(* IEC 61131-3 sources: daoli-st-library/DL_Process (part 54) *)

(* ---- FB_DL_SugarPanBatchSeq.st ---- *)
(*==============================================================================
  Component : FB_DL_SugarPanBatchSeq
  Category  : DL_Process
  Type      : FB
  Complexity: C4
  VERSION   : v1.0.0
  功能      : 煮糖罐批次时序（抽真空→进糖浆→浓缩→投晶种→助晶→终浓缩→破真空→放糖→洗罐）
  开源溯源  : 道莅原创 clean-room 自研（无外部代码引用）｜License: MIT
  边界条件  : ① 相迁移主判据为过饱和度 S（本件内联调用 CalcSupersaturation 计算）：
                 S = (Bx / (100 − Bx)) / (BxSat / (100 − BxSat))，BxSat = fSolA + fSolB × 温度；
                 该式为工程线性溶解度近似，精度受 fSolA / fSolB 标定限，不适用于高纯度精糖结晶建模。
              ② 真空与温度双联锁：真空丧失（fVacKpa 高于 fVacGoodKpa）或温度超上限 -> E3 立即断能；
                 温度低于下限 -> E2 停机待复位（糖液过冷会在罐内结块，属可恢复但需人工确认）。
              ③ 黄级语义：助晶相过饱和度超 fSWarn 只记录分级、不迁移、不置 bError（红/黑才动作）。
              ④ 过饱和度计算为「正解方向」：域外输入返回哨兵 0.0 并由调用方升 E2 上报（不静默钳位）。
                 S 物理上恒 > 1（过饱和），故 0.0 与任何合法值不重叠（R81 哨兵口径）。
                 传感器域判只在批次运行相生效——空闲相罐内空载（锤度 0、常压）属正常读数，不得误锁故障。
              ⑤ 默认引脚组合自证（R114）：握手类（bSyrupReady / bSeedAdded / bDischargeDone / bWashDone）
                 默认 FALSE，默认组合无法越过进料与放料握手直达完成相；使能类（bEStopHealthy）默认 TRUE
                 与 bEnable 同族，断线由硬件安全回路保证。
              ⑥ 复位作用域（R311）：bReset 沿清 E2/E3 锁存 + 批次计数 + 曲线锁存；bStop 只清 E2 与相位。
  状态机    : eIdle 待机 / eVacuum 抽真空 / eFillSyrup 进糖浆 / eConcentrate 浓缩到过饱和 /
              eSeed 投晶种 / eGrow 助晶养晶 / eFinalBoil 终浓缩到放糖锤度 / eBreakVac 破真空 /
              eDischarge 放糖 / eWash 洗罐 / eDone 结算拍 / eFault 停机待复位(E2) / eSafeStop 安全断能(E3)
  自检      : R1 零 GVL ｜ R2 零物理地址 ｜ R3 纯 IEC 61131-3 ｜ R4 除零先判 + 非有限自反判 ｜
              R6 CASE 含 ELSE ｜ R7 九 TON 两沿段 0 无条件刷新 ｜ R10 仅标准转换函数 ｜ R14 无属性件
==============================================================================*)
TYPE E_DL_SpbPhase :
(
    eIdle        := 0,  (* 待机：等启动沿 / Idle, waiting for start edge *)
    eVacuum      := 10, (* 抽真空相：真空度达标 / Pulling vacuum *)
    eFillSyrup   := 20, (* 进糖浆相：进料到量 / Filling syrup *)
    eConcentrate := 30, (* 浓缩相：S 到投晶目标 / Concentrating to seeding S *)
    eSeed        := 40, (* 投晶种相：晶种加入完成 / Seeding *)
    eGrow        := 50, (* 助晶相：养晶至目标 S / Crystal growing *)
    eFinalBoil   := 60, (* 终浓缩相：锤度到放糖点 / Final boil to discharge Brix *)
    eBreakVac    := 70, (* 破真空相：破真空到位 / Breaking vacuum *)
    eDischarge   := 80, (* 放糖相：放料完成 / Discharging *)
    eWash        := 90, (* 洗罐相：洗罐完成 / Pan washing *)
    eDone        := 100,(* 结算拍：批次与节拍统计 / Settlement, one-scan *)
    eFault       := 110,(* 停机待复位（E2）/ Stop awaiting reset, E2 *)
    eSafeStop    := 120 (* 安全侧断能（E3）/ Safety energy cut, E3 *)
);
END_TYPE
TYPE E_DL_SpbCause :
(
    eNone       := 0,   (* 无异常 / No anomaly *)
    eVacLost    := 1,   (* 真空度丧失（E3）/ Vacuum lost, E3 *)
    eTempHigh   := 2,   (* 罐温超上限（E3）/ Over-temperature, E3 *)
    eTempLow    := 3,   (* 罐温低于下限（E2，过冷结块）/ Under-temperature, E2 *)
    eSigBad     := 4,   (* 传感器非有限或 S 计算域外（E2）/ Non-finite signal or S out of domain, E2 *)
    eEStopOpen  := 5,   (* 急停回路断开（E3）/ E-stop open, E3 *)
    eVacTmo     := 6,   (* 抽真空超时（E2）/ Vacuum timeout, E2 *)
    eFillTmo    := 7,   (* 进糖浆超时（E2）/ Fill timeout, E2 *)
    eConcTmo    := 8,   (* 浓缩超时（E2）/ Concentrate timeout, E2 *)
    eSeedTmo    := 9,   (* 投晶种超时（E2）/ Seeding timeout, E2 *)
    eGrowTmo    := 10,  (* 助晶超时（E2）/ Growing timeout, E2 *)
    eFinalTmo   := 11,  (* 终浓缩超时（E2）/ Final boil timeout, E2 *)
    eBreakTmo   := 12,  (* 破真空超时（E2）/ Break-vacuum timeout, E2 *)
    eDischTmo   := 13,  (* 放糖超时（E2）/ Discharge timeout, E2 *)
    eWashTmo    := 14,  (* 洗罐超时（E2）/ Wash timeout, E2 *)
    eCfgBad     := 15,  (* 组态非法（E2）/ Illegal configuration, E2 *)
    ePhaseBad   := 16   (* 非法相位兜底（E2）/ Illegal phase fallback, E2 *)
);
END_TYPE
TYPE E_DL_SpbGrade :
(
    eOk     := 0,       (* 无异常 / No anomaly *)
    eYellow := 1,       (* 黄：记录并继续（S 偏离不升故障）/ Yellow, recorded only *)
    eRed    := 2,       (* 红：本批次降级（可继续至放糖）/ Red, batch degraded *)
    eBlack  := 3        (* 黑：立即断能 / Black, immediate energy cut *)
);
END_TYPE

FUNCTION_BLOCK FB_DL_SugarPanBatchSeq
VAR_INPUT
    bStart          : BOOL := FALSE;    (* 启动沿（eIdle 入 eVacuum） [-] / Start rising edge *)
    bStop           : BOOL := FALSE;    (* 中止：回 eIdle 并清 E2 锁存 [-] / Abort, clears E2 only *)
    bReset          : BOOL := FALSE;    (* 复位沿：清全部锁存 + 批次计数（R311） [-] / Reset edge *)
    bSyrupReady     : BOOL := FALSE;    (* 进糖浆到位（默认 FALSE 禁跳步） [-] / Syrup fill in position *)
    bSeedAdded      : BOOL := FALSE;    (* 晶种已加入（默认 FALSE 禁跳步） [-] / Seed added *)
    bDischargeDone  : BOOL := FALSE;    (* 放糖完成（默认 FALSE 禁跳步） [-] / Discharge done *)
    bWashDone       : BOOL := FALSE;    (* 洗罐完成（默认 FALSE 禁跳步） [-] / Wash done *)
    bEStopHealthy   : BOOL := TRUE;     (* 急停回路正常（使能类引脚，默认 TRUE） [-] / E-stop healthy *)
    fVacKpa         : LREAL := 101.3;   (* 罐内绝对压力实测（真空好 = 值低） [kPa] / Pan absolute pressure [kPa] *)
    fTempC          : LREAL := 20.0;    (* 糖液温度实测 [℃] / Syrup temperature [degC] *)
    fBrix           : LREAL := 65.0;    (* 糖液锤度实测，域 0..100 [°Bx] / Brix [degBx] *)
    fVacGoodKpa     : LREAL := 30.0;    (* 真空良好门限，域 > 0（实测 <= 该值即真空有效） [kPa] / Vacuum good limit [kPa] *)
    fTempMinC       : LREAL := 60.0;    (* 罐温下限，域 > 0（低于则 E2） [℃] / Temperature floor [degC] *)
    fTempMaxC       : LREAL := 80.0;    (* 罐温上限，域 > fTempMinC（高于则 E3） [℃] / Temperature ceiling [degC] *)
    fSolA           : LREAL := 60.0;    (* 溶解度线性式截距（标定值），域 > 0 [°Bx] / Solubility intercept [degBx] *)
    fSolB           : LREAL := 0.25;    (* 溶解度线性式斜率（标定值），域 > 0 [°Bx/℃] / Solubility slope [degBx/degC] *)
    fSSeed          : LREAL := 1.20;    (* 投晶目标过饱和度，域 > 1.0 [-] / Seeding supersaturation *)
    fSGrow          : LREAL := 1.35;    (* 助晶终点过饱和度，域 > fSSeed [-] / Growing end supersaturation *)
    fSWarn          : LREAL := 1.45;    (* 过饱和预警上界，域 > fSGrow（黄级记录） [-] / Supersaturation warn limit *)
    fBrixDischarge  : LREAL := 92.0;    (* 放糖锤度，域 0..100（且 > fBrix） [°Bx] / Discharge Brix [degBx] *)
    atPhaseTmo      : ARRAY[0..8] OF TIME := [T#20M, T#30M, T#120M, T#10M, T#240M, T#120M, T#10M, T#20M, T#30M];   (* 超时窗 [ms]，下标 0..8 = 抽真空/进料/浓缩/投晶/助晶/终浓/破真空/放糖/洗罐 / Phase windows [ms] *)
    fCycleSec       : LREAL := 0.0;     (* 扫描周期（<=0 用缺省 0.01s） [s] / Scan cycle [s] *)
END_VAR
VAR_OUTPUT
    eState          : E_DL_SpbPhase;    (* 当前相（HMI 诊断） [-] / Present phase *)
    eCause          : E_DL_SpbCause;    (* 成因（锁存回放，R189） [-] / Latched cause playback *)
    eGrade          : E_DL_SpbGrade;    (* 分级出口 [-] / Grade outlet *)
    bError          : BOOL;             (* 故障标志（E2/E3 为 TRUE） [-] / Error flag *)
    bSafeCut        : BOOL;             (* 安全侧断能指令（E3 常 TRUE 至复位） [-] / Safety energy cut *)
    bDone           : BOOL;             (* 单拍结算脉冲 [-] / One-scan done pulse *)
    bBoilActive     : BOOL;             (* 浓缩段指示（供 IO 层驱动蒸汽阀） [-] / Boiling indicator *)
    nBatchCount     : UDINT;            (* 累计批次数（饱和） [批] / Batch count, saturating *)
    fSLast          : LREAL;            (* 最近过饱和度（0 = 无效）/ 哨兵值与合法域不重叠 [-] / Last supersaturation *)
    fBrixLast       : LREAL;            (* 最近锤度 [°Bx] / Last Brix [degBx] *)
    tBatchLast      : TIME;             (* 最近一批总时长 [ms] / Last batch duration [ms] *)
END_VAR
VAR
    _ePhase      : E_DL_SpbPhase := E_DL_SpbPhase.eIdle;     (* 内部相（CASE 唯一写入目标） [-] / Internal phase *)
    _eCause      : E_DL_SpbCause := E_DL_SpbCause.eNone;     (* 成因锁存量 [-] / Latched cause *)
    _eGrade      : E_DL_SpbGrade := E_DL_SpbGrade.eOk;       (* 分级锁存量 [-] / Latched grade *)
    _bFault      : BOOL := FALSE;       (* E2 锁存位（解除 = bReset 沿或 bStop） [-] / E2 latch *)
    _bSafeLatch  : BOOL := FALSE;       (* E3 锁存位（解除 = bReset 沿且安全恢复） [-] / E3 latch *)
    _bFaultReq   : BOOL := FALSE;       (* 单拍 E2 请求（段 1 预清，段 6 落地） [-] / One-scan E2 request *)
    _bSafeReq    : BOOL := FALSE;       (* 单拍 E3 请求（段 1 预清，段 6 落地） [-] / One-scan E3 request *)
    _bDonePulse  : BOOL := FALSE;       (* 单拍结算标志（段 1 预清） [-] / One-scan done flag *)
    _bVacOk      : BOOL := FALSE;       (* 真空有效判据 [-] / Vacuum valid *)
    _bTempHigh   : BOOL := FALSE;       (* 罐温超上限当拍量 [-] / Over-temperature this scan *)
    _bTempLow    : BOOL := FALSE;       (* 罐温低于下限当拍量 [-] / Under-temperature this scan *)
    _bVacBad     : BOOL := FALSE;       (* 真空传感器非有限当拍量 [-] / Vacuum non-finite *)
    _bTempBad    : BOOL := FALSE;       (* 温度传感器非有限当拍量 [-] / Temperature non-finite *)
    _bBrixBad    : BOOL := FALSE;       (* 锤度非有限或域外当拍量 [-] / Brix non-finite or out of domain *)
    _bCfgBad     : BOOL := FALSE;       (* 组态非法当拍量 [-] / Configuration bad *)
    _fS          : LREAL := 0.0;        (* 当拍过饱和度（0 = 计算无效哨兵） [-] / Supersaturation this scan *)
    _fMsTmp      : LREAL := 0.0;        (* 批次时长毫秒暂存（转换前钳位） [ms] / Batch milliseconds scratch *)
    _bVacRequired: BOOL := FALSE;       (* 本相要求真空有效（进料至终浓缩）/ Vacuum required in phase *)
    _bBatchActive: BOOL := FALSE;       (* 批次运行相（空闲与故障相不计信号域判）/ Batch active phase *)
    _bSafeOk     : BOOL := FALSE;       (* 安全条件已恢复（E3 解除判据）/ Safety conditions recovered *)
    _fBrixLatch  : LREAL := 0.0;        (* 锤度锁存（出口留影） [°Bx] / Brix latch *)
    _fBatchAccS  : LREAL := 0.0;        (* 本批时长累加 [s] / Batch time accumulator *)
    _tBatchLast  : TIME := T#0S;        (* 最近批时长锁存 [ms] / Last batch duration latch *)
    _fCy         : LREAL := 0.0;        (* 当拍有效周期 [s] / Effective cycle *)
    _nBatch      : UDINT := 0;          (* 批次累计锁存（饱和） [批] / Batch count latch *)
    _nIdxChk     : INT := 0;            (* 相窗遍历索引（循环变量） [-] / Loop index *)
    tonVacuum    : TON;                 (* 抽真空超时（段 0 无条件调用） / Vacuum timeout *)
    tonFill      : TON;                 (* 进糖浆超时 / Fill timeout *)
    tonConcentrate: TON;                (* 浓缩超时 / Concentrate timeout *)
    tonSeed      : TON;                 (* 投晶种超时 / Seeding timeout *)
    tonGrow      : TON;                 (* 助晶超时 / Growing timeout *)
    tonFinalBoil : TON;                 (* 终浓缩超时 / Final boil timeout *)
    tonBreakVac  : TON;                 (* 破真空超时 / Break-vacuum timeout *)
    tonDischarge : TON;                 (* 放糖超时 / Discharge timeout *)
    tonWash      : TON;                 (* 洗罐超时 / Wash timeout *)
    rtStart      : R_TRIG;              (* 启动沿（段 0 无条件调用） / Start edge *)
    rtReset      : R_TRIG;              (* 复位沿（段 0 无条件调用） / Reset edge *)
END_VAR
VAR CONSTANT
    DL_SPB_CYDEF   : LREAL := 0.01;         (* 缺省扫描周期 [s] / Default scan cycle [s] *)
    DL_SPB_BRIXTOP : LREAL := 100.0;        (* 锤度与溶解度共用上界 [°Bx] / Brix and solubility ceiling *)
    DL_SPB_DENMIN  : LREAL := 1.0E-6;       (* 除法分母下限（判零） [-] / Divisor floor *)
    DL_SPB_BATMAX  : UDINT := 4294967295;   (* 批次计数饱和上限 [批] / Batch count ceiling *)
END_VAR

(*-----------------------------------------------------------------------------
  方法 CalcSupersaturation：过饱和度计算（正解方向，域闸四段式）
  四段：① 返回值预置哨兵 0.0 ② 域闸命中直接 RETURN（非有限 / 锤度域外 / 溶解度域外）
        ③ 域内才做两次除法（分母均已证明 > DL_SPB_DENMIN） ④ 结果非有限复检兜底
  契约：返回 0.0 = 计算无效（哨兵），S 物理恒 > 1，调用方据 0.0 升 E2 上报（禁静默钳位）。
-----------------------------------------------------------------------------*)
METHOD PUBLIC CalcSupersaturation : LREAL
VAR_INPUT
    fBrixIn  : LREAL := 0.0;    (* 锤度输入，域 (0, 100) [°Bx] / Brix input *)
    fTempIn  : LREAL := 0.0;    (* 温度输入 [℃] / Temperature input *)
    fSolAIn  : LREAL := 0.0;    (* 溶解度截距，域 > 0 [°Bx] / Solubility intercept *)
    fSolBIn  : LREAL := 0.0;    (* 溶解度斜率，域 > 0 [°Bx/℃] / Solubility slope *)
END_VAR
VAR
    fBxSat : LREAL := 0.0;      (* 该温度下饱和锤度 [°Bx] / Saturated Brix at temperature *)
    fNum   : LREAL := 0.0;      (* 分子 Bx / (100 − Bx) [-] / Numerator *)
    fDen   : LREAL := 0.0;      (* 分母 BxSat / (100 − BxSat) [-] / Denominator *)
    fS     : LREAL := 0.0;      (* 过饱和度暂存 [-] / Supersaturation scratch *)
END_VAR

CalcSupersaturation := 0.0;     (* ① 预置哨兵 / Preset sentinel *)
IF (fBrixIn <> fBrixIn) OR ((fBrixIn - fBrixIn) <> (fBrixIn - fBrixIn)) THEN
    CalcSupersaturation := 0.0; (* ② 锤度非有限 / Brix non-finite *)
    RETURN;
END_IF
IF (fTempIn <> fTempIn) OR ((fTempIn - fTempIn) <> (fTempIn - fTempIn)) THEN
    CalcSupersaturation := 0.0; (* ② 温度非有限 / Temperature non-finite *)
    RETURN;
END_IF
IF (fSolAIn <= 0.0) OR (fSolBIn <= 0.0) THEN
    CalcSupersaturation := 0.0; (* ② 溶解度系数域外 / Solubility coefficient out of domain *)
    RETURN;
END_IF
IF (fBrixIn <= 0.0) OR (fBrixIn >= DL_SPB_BRIXTOP) THEN
    CalcSupersaturation := 0.0; (* ② 锤度域外（分母 100 − Bx 失效保护）/ Brix out of domain *)
    RETURN;
END_IF
fBxSat := fSolAIn + fSolBIn * fTempIn;                         (* 线性溶解度式 [°Bx] / Linear solubility *)
IF (fBxSat <= 0.0) OR (fBxSat >= DL_SPB_BRIXTOP) THEN
    CalcSupersaturation := 0.0; (* ② 饱和锤度域外 / Saturated Brix out of domain *)
    RETURN;
END_IF
fNum := fBrixIn / (DL_SPB_BRIXTOP - fBrixIn);                   (* ③ 分母 > 0 已证 / Denominator proven positive *)
fDen := fBxSat / (DL_SPB_BRIXTOP - fBxSat);                     (* ③ 分母 > 0 已证 / Denominator proven positive *)
IF fDen < DL_SPB_DENMIN THEN
    CalcSupersaturation := 0.0; (* ③ 分母判零（防御式，域闸后不可达）/ Divisor guard *)
    RETURN;
END_IF
fS := fNum / fDen;                                             (* 过饱和度 [-] / Supersaturation *)
IF (fS <> fS) OR ((fS - fS) <> (fS - fS)) THEN
    CalcSupersaturation := 0.0; (* ④ 结果非有限兜底 / Result non-finite fallback *)
    RETURN;
END_IF
CalcSupersaturation := fS;                                     (* 合法结果输出 / Valid result *)
END_METHOD

(*-----------------------------------------------------------------------------
  方法 ResetBatch：批次锁存复位（不清累计批次数，累计量只能由 bReset 沿清除）
  契约：返回 TRUE 表示复位执行；作用于分级、成因、过饱和度锁存与批次时长累加。
-----------------------------------------------------------------------------*)
METHOD PUBLIC ResetBatch : BOOL
ResetBatch := FALSE;                            (* 预置 / Preset *)
_eGrade := E_DL_SpbGrade.eOk;                   (* 清分级 / Clear grade *)
_eCause := E_DL_SpbCause.eNone;                 (* 清成因 / Clear cause *)
_fS := 0.0;                                     (* 清过饱和度哨兵 / Clear supersaturation *)
_fBrixLatch := 0.0;                             (* 清锤度锁存 / Clear Brix latch *)
_fBatchAccS := 0.0;                             (* 清批次时长累加 / Clear batch accumulator *)
ResetBatch := TRUE;                             (* 复位已执行 / Reset performed *)
END_METHOD

(* —— 段 0：传感器非有限与域判 + 过饱和度计算 + 组态闸 + 周期 + 九 TON 两沿无条件刷新（R7） —— *)
_bVacBad := (fVacKpa <> fVacKpa) OR ((fVacKpa - fVacKpa) <> (fVacKpa - fVacKpa));      (* NaN 自反 + Inf 差值 / NaN and Inf *)
_bTempBad := (fTempC <> fTempC) OR ((fTempC - fTempC) <> (fTempC - fTempC));
_bBrixBad := (fBrix <> fBrix) OR ((fBrix - fBrix) <> (fBrix - fBrix))
          OR (fBrix <= 0.0) OR (fBrix >= DL_SPB_BRIXTOP);                             (* 锤度域外并入信号级 / Brix domain *)
_bVacOk := (NOT _bVacBad) AND (fVacKpa <= fVacGoodKpa);                                (* 真空有效（值低为好）/ Vacuum valid *)
_bTempHigh := (NOT _bTempBad) AND (fTempC > fTempMaxC);                                (* 超上限（E3）/ Over-temperature *)
_bTempLow := (NOT _bTempBad) AND (fTempC < fTempMinC);                                 (* 低于下限（E2）/ Under-temperature *)
_fS := CalcSupersaturation(fBrix, fTempC, fSolA, fSolB);                               (* 过饱和度内联计算 / Supersaturation *)
_bCfgBad := (fVacGoodKpa <= 0.0) OR (fTempMinC <= 0.0) OR (fTempMaxC <= fTempMinC)
         OR (fSolA <= 0.0) OR (fSolB <= 0.0) OR (fBrixDischarge <= 0.0)
         OR (fBrixDischarge >= DL_SPB_BRIXTOP) OR (fSSeed <= 1.0)
         OR (fSGrow <= fSSeed) OR (fSWarn <= fSGrow);                                 (* 组态域闸与配比 / Config gate *)
FOR _nIdxChk := 0 TO 8 DO
    IF atPhaseTmo[_nIdxChk] <= T#0S THEN
        _bCfgBad := TRUE;                                                             (* 任一相窗非正 -> 组态非法 / Non-positive window *)
    END_IF
END_FOR
IF fCycleSec > 0.0 THEN
    _fCy := fCycleSec;                                                                (* 组态周期有效 / Configured cycle *)
ELSE
    _fCy := DL_SPB_CYDEF;                                                             (* 周期缺省兜底 / Default cycle *)
END_IF
rtStart(CLK := bStart);                                                               (* 启动沿，每拍必调 / Start edge every scan *)
rtReset(CLK := bReset);                                                               (* 复位沿，每拍必调 / Reset edge every scan *)
tonVacuum(IN := (_ePhase = E_DL_SpbPhase.eVacuum), PT := atPhaseTmo[0]);              (* 抽真空窗 / Vacuum window *)
tonFill(IN := (_ePhase = E_DL_SpbPhase.eFillSyrup), PT := atPhaseTmo[1]);             (* 进料窗 / Fill window *)
tonConcentrate(IN := (_ePhase = E_DL_SpbPhase.eConcentrate), PT := atPhaseTmo[2]);    (* 浓缩窗 / Concentrate window *)
tonSeed(IN := (_ePhase = E_DL_SpbPhase.eSeed), PT := atPhaseTmo[3]);                  (* 投晶窗 / Seeding window *)
tonGrow(IN := (_ePhase = E_DL_SpbPhase.eGrow), PT := atPhaseTmo[4]);                  (* 助晶窗 / Growing window *)
tonFinalBoil(IN := (_ePhase = E_DL_SpbPhase.eFinalBoil), PT := atPhaseTmo[5]);        (* 终浓窗 / Final boil window *)
tonBreakVac(IN := (_ePhase = E_DL_SpbPhase.eBreakVac), PT := atPhaseTmo[6]);          (* 破真空窗 / Break vacuum window *)
tonDischarge(IN := (_ePhase = E_DL_SpbPhase.eDischarge), PT := atPhaseTmo[7]);        (* 放糖窗 / Discharge window *)
tonWash(IN := (_ePhase = E_DL_SpbPhase.eWash), PT := atPhaseTmo[8]);                  (* 洗罐窗 / Wash window *)

(* —— 段 1：单拍量预清零（不含锁存/累加/计数，R107）+ 批次时长累加 —— *)
_bFaultReq := FALSE;                                                                  (* E2 请求预清 / E2 request preset *)
_bSafeReq := FALSE;                                                                   (* E3 请求预清 / E3 request preset *)
_bDonePulse := FALSE;                                                                 (* 结算标志预清 / Done preset *)
bError := FALSE;                                                                      (* 故障标志预清（出口汇总）/ Error preset *)
IF (_ePhase <> E_DL_SpbPhase.eIdle) AND (_ePhase <> E_DL_SpbPhase.eFault)
   AND (_ePhase <> E_DL_SpbPhase.eSafeStop) THEN
    _fBatchAccS := _fBatchAccS + _fCy;                                                (* 批次时长累加（仅工作相）/ Batch time, working phases only *)
END_IF
_bVacRequired := (_ePhase = E_DL_SpbPhase.eFillSyrup) OR (_ePhase = E_DL_SpbPhase.eConcentrate)
              OR (_ePhase = E_DL_SpbPhase.eSeed) OR (_ePhase = E_DL_SpbPhase.eGrow)
              OR (_ePhase = E_DL_SpbPhase.eFinalBoil);                                (* 真空维持段（放糖与洗罐不要求）/ Vacuum-required phases *)
_bBatchActive := (_ePhase <> E_DL_SpbPhase.eIdle) AND (_ePhase <> E_DL_SpbPhase.eDone)
                   AND (_ePhase <> E_DL_SpbPhase.eVacuum) AND (_ePhase <> E_DL_SpbPhase.eFillSyrup)   (* 空罐与进料相锤度天然为 0，不计入信号域判 / Exclude vacuum & fill phases: brix is naturally 0 *)
              AND (_ePhase <> E_DL_SpbPhase.eFault) AND (_ePhase <> E_DL_SpbPhase.eSafeStop);   (* 批次运行相判据 / Batch-active judge *)
_bSafeOk := bEStopHealthy AND (NOT _bTempHigh) AND (NOT _bTempBad);                   (* 安全恢复基础判据 / Base safety recovery *)
IF _eCause = E_DL_SpbCause.eVacLost THEN
    _bSafeOk := _bSafeOk AND _bVacOk;                                                 (* 真空成因须真空恢复（R152 可达性）/ Vacuum cause needs vacuum back *)
END_IF

(* —— 段 2：E3 安全侧（急停 / 真空丧失 / 罐温超上限）——最高优先级 —— *)
IF NOT bEStopHealthy THEN
    IF NOT _bSafeLatch THEN
        _bSafeReq := TRUE;                                                            (* 落地于段 6 / Landed in segment 6 *)
        _eCause := E_DL_SpbCause.eEStopOpen;                                          (* 归因：急停断开 / Cause: E-stop *)
    END_IF
ELSIF _bTempHigh THEN
    IF NOT _bSafeLatch THEN
        _bSafeReq := TRUE;
        _eCause := E_DL_SpbCause.eTempHigh;                                           (* 归因：超温 / Cause: over-temperature *)
    END_IF
ELSIF _bVacRequired AND (NOT _bVacBad) AND (NOT _bVacOk) THEN
    IF NOT _bSafeLatch THEN
        _bSafeReq := TRUE;                                                            (* 真空在非抽真空相丧失：立即断能 / Vacuum lost mid-batch *)
        _eCause := E_DL_SpbCause.eVacLost;                                            (* 归因：真空丧失 / Cause: vacuum lost *)
    END_IF
END_IF

(* —— 段 3：信号域闸与组态闸入 E2（E3 优先，安全相内不重复置因） —— *)
IF _bCfgBad AND (NOT _bSafeLatch) AND (NOT _bFault) THEN
    _bFaultReq := TRUE;                                                               (* 落地于段 6 / Landed in segment 6 *)
    _eCause := E_DL_SpbCause.eCfgBad;                                                 (* 归因：组态非法 / Cause: config *)
ELSIF _bBatchActive AND (_bVacBad OR _bBrixBad) THEN
    IF NOT _bSafeLatch AND NOT _bFault THEN
        _bFaultReq := TRUE;
        _eCause := E_DL_SpbCause.eSigBad;                                             (* 归因：传感器非有限 / Cause: non-finite *)
    END_IF
ELSIF _bBatchActive AND _bTempLow THEN
    IF NOT _bSafeLatch AND NOT _bFault THEN
        _bFaultReq := TRUE;
        _eCause := E_DL_SpbCause.eTempLow;                                            (* 归因：过冷 / Cause: under-temperature *)
    END_IF
ELSIF _bBatchActive AND (_fS <= 0.0) AND (NOT _bFault) THEN
    IF NOT _bSafeLatch THEN
        _bFaultReq := TRUE;                                                           (* S 计算域外（哨兵 0.0）/ S sentinel zero *)
        _eCause := E_DL_SpbCause.eSigBad;                                             (* 归因：S 计算域外 / Cause: S out of domain *)
    END_IF
END_IF

(* —— 段 4：迁出链（复位沿 > 中止；作用域逐项声明 R311） —— *)
IF rtReset.Q THEN
    _bFault := FALSE;                                                                 (* 作用域①：清 E2 锁存 / Clear E2 *)
    IF _bSafeOk THEN
        _bSafeLatch := FALSE;                                                         (* 作用域②：安全恢复才清 E3（成因相关判据）/ Clear E3 only if safe *)
    END_IF
    _eCause := E_DL_SpbCause.eNone;                                                   (* 作用域③：清成因分级 / Clear cause and grade *)
    _eGrade := E_DL_SpbGrade.eOk;
    _fS := 0.0;                                                                       (* 作用域④：清过饱和度锁存 / Clear supersaturation *)
    _fBrixLatch := 0.0;
    _fBatchAccS := 0.0;                                                               (* 作用域⑤：清批次时长 / Clear batch time *)
    _nBatch := 0;                                                                     (* 作用域⑥：清批次计数（生产资料复位）/ Clear batch count *)
    IF NOT _bSafeLatch THEN
        IF (_ePhase = E_DL_SpbPhase.eFault) OR (_ePhase = E_DL_SpbPhase.eSafeStop) THEN
            _ePhase := E_DL_SpbPhase.eIdle;                                           (* 作用域⑦：故障相迁回待机 / Back to idle *)
        END_IF
    END_IF
ELSIF bStop AND (_ePhase <> E_DL_SpbPhase.eIdle) AND (_ePhase <> E_DL_SpbPhase.eSafeStop) THEN
    IF _ePhase = E_DL_SpbPhase.eFault THEN
        _bFault := FALSE;                                                             (* 中止清 E2（E3 只由复位清）/ Abort clears E2 only *)
        _eCause := E_DL_SpbCause.eNone;
        _eGrade := E_DL_SpbGrade.eOk;
    END_IF
    _fBatchAccS := 0.0;                                                               (* 批次时长作废 / Batch time void *)
    _ePhase := E_DL_SpbPhase.eIdle;                                                   (* 回待机 / Back to idle *)
END_IF

(* —— 段 5：主状态机（过饱和度 / 锤度为相迁移主判据，超时为保护） —— *)
CASE _ePhase OF
E_DL_SpbPhase.eIdle:
    IF rtStart.Q AND (NOT _bFault) AND (NOT _bSafeLatch) THEN
        _eGrade := E_DL_SpbGrade.eOk;                                                 (* 新批起算 / New batch *)
        _eCause := E_DL_SpbCause.eNone;
        _fBatchAccS := 0.0;
        _ePhase := E_DL_SpbPhase.eVacuum;                                             (* 入抽真空相 / To vacuum *)
    END_IF
E_DL_SpbPhase.eVacuum:
    IF _bVacOk THEN
        _ePhase := E_DL_SpbPhase.eFillSyrup;                                          (* 真空达标 -> 进糖浆 / Vacuum OK, fill *)
    ELSIF tonVacuum.Q THEN
        _eCause := E_DL_SpbCause.eVacTmo;                                             (* 归因：抽真空超时 / Cause: vacuum timeout *)
        _bFaultReq := TRUE;
    END_IF
E_DL_SpbPhase.eFillSyrup:
    IF bSyrupReady THEN
        _ePhase := E_DL_SpbPhase.eConcentrate;                                        (* 进料到量 -> 浓缩 / Filled, concentrate *)
    ELSIF tonFill.Q THEN
        _eCause := E_DL_SpbCause.eFillTmo;                                            (* 归因：进料超时 / Cause: fill timeout *)
        _bFaultReq := TRUE;
    END_IF
E_DL_SpbPhase.eConcentrate:
    IF (_fS > 0.0) AND (_fS >= fSSeed) THEN
        _ePhase := E_DL_SpbPhase.eSeed;                                               (* S 到投晶目标 -> 投晶 / S reached, seed *)
    ELSIF tonConcentrate.Q THEN
        _eCause := E_DL_SpbCause.eConcTmo;                                            (* 归因：浓缩超时（S 未达）/ Cause: concentrate timeout *)
        _bFaultReq := TRUE;
    END_IF
E_DL_SpbPhase.eSeed:
    IF bSeedAdded THEN
        _ePhase := E_DL_SpbPhase.eGrow;                                               (* 晶种加入 -> 助晶 / Seeded, grow *)
    ELSIF tonSeed.Q THEN
        _eCause := E_DL_SpbCause.eSeedTmo;                                            (* 归因：投晶超时 / Cause: seeding timeout *)
        _bFaultReq := TRUE;
    END_IF
E_DL_SpbPhase.eGrow:
    IF (_fS > 0.0) AND (_fS > fSWarn) THEN
        _eGrade := E_DL_SpbGrade.eYellow;                                             (* 过饱和偏高预警（黄，只记录不迁移）/ High-S warning, recorded only *)
    END_IF
    IF (_fS > 0.0) AND (_fS >= fSGrow) THEN
        _ePhase := E_DL_SpbPhase.eFinalBoil;                                          (* 养晶到位 -> 终浓 / Grown, final boil *)
    ELSIF tonGrow.Q THEN
        _eCause := E_DL_SpbCause.eGrowTmo;                                            (* 归因：助晶超时 / Cause: growing timeout *)
        _bFaultReq := TRUE;
    END_IF
E_DL_SpbPhase.eFinalBoil:
    IF (NOT _bBrixBad) AND (fBrix >= fBrixDischarge) THEN
        _fBrixLatch := fBrix;                                                         (* 放糖锤度锁存 / Latch discharge Brix *)
        _ePhase := E_DL_SpbPhase.eBreakVac;                                           (* 锤度到量 -> 破真空 / Brix reached, break vacuum *)
    ELSIF tonFinalBoil.Q THEN
        _eCause := E_DL_SpbCause.eFinalTmo;                                           (* 归因：终浓超时（锤度未达）/ Cause: final boil timeout *)
        _bFaultReq := TRUE;
    END_IF
E_DL_SpbPhase.eBreakVac:
    IF (NOT _bVacBad) AND (fVacKpa >= fVacGoodKpa) THEN
        _ePhase := E_DL_SpbPhase.eDischarge;                                          (* 真空破除到位 -> 放糖（本拍事件优先，R275）/ Vacuum broken, discharge *)
    ELSIF tonBreakVac.Q THEN
        _eCause := E_DL_SpbCause.eBreakTmo;                                           (* 归因：破真空超时 / Cause: break-vacuum timeout *)
        _bFaultReq := TRUE;
    END_IF
E_DL_SpbPhase.eDischarge:
    IF bDischargeDone THEN
        _ePhase := E_DL_SpbPhase.eWash;                                               (* 放糖完成 -> 洗罐 / Discharged, wash *)
    ELSIF tonDischarge.Q THEN
        _eCause := E_DL_SpbCause.eDischTmo;                                           (* 归因：放糖超时 / Cause: discharge timeout *)
        _bFaultReq := TRUE;
    END_IF
E_DL_SpbPhase.eWash:
    IF bWashDone THEN
        _ePhase := E_DL_SpbPhase.eDone;                                               (* 洗罐完成 -> 结算 / Washed, settle *)
    ELSIF tonWash.Q THEN
        _eCause := E_DL_SpbCause.eWashTmo;                                            (* 归因：洗罐超时 / Cause: wash timeout *)
        _bFaultReq := TRUE;
    END_IF
E_DL_SpbPhase.eDone:
    _bDonePulse := TRUE;                                                              (* 单拍结算（段 1 预清）/ One-scan done *)
    _fMsTmp := _fBatchAccS * 1000.0;                                                  (* 秒 -> 毫秒 [ms] / Second to millisecond *)
    IF _fMsTmp > 2147483647.0 THEN
        _fMsTmp := 2147483647.0;                                                      (* 取整前实数上限兜底（R153）/ Real ceiling before truncation *)
    END_IF
    _tBatchLast := DINT_TO_TIME(LREAL_TO_DINT(_fMsTmp));                              (* 批次时长换算 / Batch duration *)
    _fBatchAccS := 0.0;                                                               (* 累加清零 / Clear accumulator *)
    IF _nBatch < DL_SPB_BATMAX THEN
        _nBatch := _nBatch + 1;                                                       (* 批次推进（容量载体判上限）/ Saturating batch count *)
    END_IF
    _ePhase := E_DL_SpbPhase.eIdle;                                                   (* 回待机 / Back to idle *)
E_DL_SpbPhase.eFault:
    bError := TRUE;                                                                   (* 故障相驻留（锁存回放）/ Fault residency *)
E_DL_SpbPhase.eSafeStop:
    bError := TRUE;                                                                   (* 安全相驻留（锁存回放）/ Safety residency *)
ELSE
    _eCause := E_DL_SpbCause.ePhaseBad;                                               (* 非法相位兜底 / Illegal phase fallback *)
    _bFaultReq := TRUE;                                                               (* 由段 6 落地 / Landed in segment 6 *)
END_CASE

(* —— 段 6：E2/E3 请求统一落地（分支内只写成因与请求，落地仅此一处，R187/R252） —— *)
IF _bSafeReq AND (NOT _bSafeLatch) THEN
    _bSafeLatch := TRUE;                                                              (* E3 锁存 / Latch E3 *)
    _eGrade := E_DL_SpbGrade.eBlack;                                                  (* 分级黑 / Grade black *)
    _ePhase := E_DL_SpbPhase.eSafeStop;                                               (* 同步迁相 / Migrate *)
    bError := TRUE;                                                                   (* 故障标志同段置位（R45 配对）/ Error pairing *)
ELSIF _bFaultReq AND (NOT _bSafeLatch) THEN
    _bFault := TRUE;                                                                  (* E2 锁存 / Latch E2 *)
    _eGrade := E_DL_SpbGrade.eRed;                                                    (* 分级红（批次降级）/ Grade red *)
    _ePhase := E_DL_SpbPhase.eFault;                                                  (* 同步迁相（R252）/ Migrate *)
    bError := TRUE;                                                                   (* 故障标志同段置位（R45 配对）/ Error pairing *)
END_IF

(* —— 段 7：统一出口（电平量由 _ePhase 派生，连续量做有限性防护 R273） —— *)
eState := _ePhase;                                                                    (* 相出口 / Phase outlet *)
eCause := _eCause;                                                                    (* 成因回放 / Cause playback *)
eGrade := _eGrade;                                                                    (* 分级出口 / Grade outlet *)
bError := bError OR _bFault OR _bSafeLatch;                                           (* 故障标志汇总 / Error summary *)
bSafeCut := _bSafeLatch;                                                              (* 安全断能指令 / Safety energy cut *)
bDone := _bDonePulse;                                                                 (* 单拍结算脉冲 / One-scan done *)
bBoilActive := (_ePhase = E_DL_SpbPhase.eConcentrate) OR (_ePhase = E_DL_SpbPhase.eGrow)
            OR (_ePhase = E_DL_SpbPhase.eFinalBoil);                                  (* 浓缩段指示 / Boiling indicator *)
nBatchCount := _nBatch;                                                               (* 批次计数出口 / Batch count outlet *)
IF (_fS <> _fS) OR ((_fS - _fS) <> (_fS - _fS)) THEN
    fSLast := 0.0;                                                                    (* 非有限不出口（保持哨兵）/ Non-finite not exported *)
ELSE
    fSLast := _fS;                                                                    (* 过饱和度出口 / Supersaturation outlet *)
END_IF
IF (_fBrixLatch <> _fBrixLatch) OR ((_fBrixLatch - _fBrixLatch) <> (_fBrixLatch - _fBrixLatch)) THEN
    fBrixLast := 0.0;                                                                 (* 非有限不出口 / Non-finite not exported *)
ELSE
    fBrixLast := _fBrixLatch;                                                         (* 锤度出口 / Brix outlet *)
END_IF
tBatchLast := _tBatchLast;                                                            (* 批次时长出口 [ms] / Batch duration outlet *)
END_FUNCTION_BLOCK

(* ---- FB_DL_TabletCompactionSeq.st ---- *)
(*
  DL Factory R84 | FB_DL_TabletCompactionSeq
  功能：压片七相时序状态机，含预压/主压到位超时、剔废计数与完成脉冲
  开源溯源：无（clean-room 自研，依据公开工艺公式，来源=行业通用公式，许可证=MIT，借鉴点=公式结构）
  规则：R1-R16 全遵守
*)
TYPE E_DL_TabCompState :
(
    eIdle := 0, // 空闲待启动 [-] / idle [-]
    eFill := 1, // 充填相 [-] / die filling phase [-]
    ePreComp := 2, // 预压相 [-] / pre compaction phase [-]
    eMainComp := 3, // 主压相 [-] / main compaction phase [-]
    eEject := 4, // 出片相 [-] / ejection phase [-]
    eRejectCheck := 5, // 剔废判定相 [-] / reject check phase [-]
    eDone := 6, // 完成相 [-] / done phase [-]
    eFault := 7 // 故障锁存相 [-] / fault latched phase [-]
) := eIdle;
END_TYPE

FUNCTION_BLOCK FB_DL_TabletCompactionSeq
VAR_INPUT
    xStart : BOOL; // 压片启动按钮 [-] / start pushbutton [-]
    xReset : BOOL; // 复位按钮，上升沿清故障码 [-] / reset pushbutton [-]
    xFillDone : BOOL; // 充填到位反馈 [-] / fill complete feedback [-]
    xPrePressOk : BOOL; // 预压压力到位反馈 [-] / pre compaction pressure reached [-]
    xMainPressOk : BOOL; // 主压压力到位反馈 [-] / main compaction pressure reached [-]
    xEjectDone : BOOL; // 出片到位反馈 [-] / ejection complete feedback [-]
    xPartOk : BOOL; // 剔废检测判定（TRUE=合格） [-] / tablet quality verdict [-]
    tFillLimit : TIME := T#5S; // 充填相超时 [s] / fill phase timeout [s]
    tEjectLimit : TIME := T#5S; // 出片相超时（独立整定，R572） [s] / eject phase timeout, tuned separately [s]
    tPreLimit : TIME := T#3S; // 预压到位超时 [s] / pre compaction timeout [s]
    tMainLimit : TIME := T#5S; // 主压到位超时 [s] / main compaction timeout [s]
END_VAR
VAR_OUTPUT
    eState : E_DL_TabCompState; // 当前时序状态 [-] / current sequence state [-]
    iErrCode : INT; // 故障码 0=正常，401~405 [-] / error code, 401 to 405 [code]
    iRejectCnt : INT; // 剔废累计片数 [片] / rejected tablet counter [tablets]
    xDone : BOOL; // 完成单拍脉冲 [-] / done one-shot pulse [-]
END_VAR
VAR
    rtStart : R_TRIG; // 启动上升沿实例 [-] / start rising edge instance [-]
    rtReset : R_TRIG; // 复位上升沿实例 [-] / reset rising edge instance [-]
    tonFill : TON; // 充填相超时定时器（独立，R572） [-] / fill phase timer, dedicated [-]
    tonEject : TON; // 出片相超时定时器（独立，R572） [-] / eject phase timer, dedicated [-]
    tonPre : TON; // 预压到位超时定时器 [-] / pre compaction timer [-]
    tonMain : TON; // 主压到位超时定时器 [-] / main compaction timer [-]
    _eState : E_DL_TabCompState := E_DL_TabCompState.eIdle; // 内部相位（CASE 唯一写目标） [-] / internal phase [-]
    _iErr : INT; // 故障码内部锁存 [-] / latched error code [-]
    _iRej : INT; // 剔废计数内部量 [片] / internal reject counter [tablets]
    xDoneInt : BOOL; // 完成内部锁存位 [-] / internal done latch [-]
    xDonePrev : BOOL; // 完成前拍快照 [-] / done previous scan snapshot [-]
END_VAR

// 段 0｜边沿与定时器实例无条件周期刷新（R7；相闸串在 IN 上）
rtStart(CLK := xStart); // 启动沿每拍必调 [-] / start edge every scan [-]
rtReset(CLK := xReset); // 复位沿每拍必调 [-] / reset edge every scan [-]
tonFill(IN := _eState = E_DL_TabCompState.eFill, PT := tFillLimit); // 充填相独立闸，离相复位 [-] / fill phase gate, reset when the phase leaves [-]
tonEject(IN := _eState = E_DL_TabCompState.eEject, PT := tEjectLimit); // 出片相独立闸，离相复位 [-] / eject phase gate, reset when the phase leaves [-]
tonPre(IN := _eState = E_DL_TabCompState.ePreComp, PT := tPreLimit); // 预压相闸 [-] / pre compaction phase gate [-]
tonMain(IN := _eState = E_DL_TabCompState.eMainComp, PT := tMainLimit); // 主压相闸 [-] / main compaction phase gate [-]

// 段 1｜复位沿：清故障码与相位（剔废计数属工艺累计量，不随复位清零，R189）
IF rtReset.Q THEN
    _iErr := 0; // 清故障码 [-] / clear error code [-]
    xDoneInt := FALSE; // 清完成锁存 [-] / clear done latch [-]
    _eState := E_DL_TabCompState.eIdle; // 回空闲相 [-] / back to idle [-]
END_IF

// 段 2｜主状态机（合法事件优先于超时迁移，R275）
CASE _eState OF
    E_DL_TabCompState.eIdle: // 空闲相 [-] / idle [-]
        xDoneInt := FALSE; // 空闲清完成锁存 [-] / clear done latch in idle [-]
        IF rtStart.Q THEN
            _eState := E_DL_TabCompState.eFill; // 启动沿进充填相 [-] / start edge enters filling [-]
        END_IF
    E_DL_TabCompState.eFill: // 充填相 [-] / filling [-]
        IF xFillDone AND NOT tonFill.Q THEN
            _eState := E_DL_TabCompState.ePreComp; // 充填到位转预压 [-] / fill done leads to pre compaction [-]
        ELSIF tonFill.Q THEN
            _iErr := 401; _eState := E_DL_TabCompState.eFault; // 充填超时（料斗缺料/下料不畅） [-] / fill timeout [-]
        END_IF
    E_DL_TabCompState.ePreComp: // 预压相 [-] / pre compaction [-]
        IF xPrePressOk AND NOT tonPre.Q THEN
            _eState := E_DL_TabCompState.eMainComp; // 预压到位转主压 [-] / pre pressure reached leads to main compaction [-]
        ELSIF tonPre.Q THEN
            _iErr := 402; _eState := E_DL_TabCompState.eFault; // 预压到位超时 [-] / pre compaction timeout [-]
        END_IF
    E_DL_TabCompState.eMainComp: // 主压相 [-] / main compaction [-]
        IF xMainPressOk AND NOT tonMain.Q THEN
            _eState := E_DL_TabCompState.eEject; // 主压到位转出片 [-] / main pressure reached leads to ejection [-]
        ELSIF tonMain.Q THEN
            _iErr := 403; _eState := E_DL_TabCompState.eFault; // 主压到位超时（液压/过载） [-] / main compaction timeout [-]
        END_IF
    E_DL_TabCompState.eEject: // 出片相 [-] / ejection [-]
        IF xEjectDone AND NOT tonEject.Q THEN
            _eState := E_DL_TabCompState.eRejectCheck; // 出片到位转剔废判定 [-] / ejection leads to reject check [-]
        ELSIF tonEject.Q THEN
            _iErr := 404; _eState := E_DL_TabCompState.eFault; // 出片到位超时 [-] / ejection timeout [-]
        END_IF
    E_DL_TabCompState.eRejectCheck: // 剔废判定相 [-] / reject check [-]
        IF xPartOk THEN
            _eState := E_DL_TabCompState.eDone; // 判定合格转完成相 [-] / qualified leads to done [-]
        ELSE
            _iRej := _iRej + 1; // 片数累加（+1 片） / count one rejected tablet
            _eState := E_DL_TabCompState.eDone; // 判废踢出后同样回完成相 [-] / rejected tablet still ends the cycle [-]
        END_IF
    E_DL_TabCompState.eDone: // 完成相 [-] / done [-]
        xDoneInt := TRUE; // 置完成锁存（出口统一映射单拍） [-] / raise done latch [-]
        IF NOT xStart THEN
            _eState := E_DL_TabCompState.eIdle; // 松开启动即回空闲 [-] / start released returns to idle [-]
        END_IF
    E_DL_TabCompState.eFault: // 故障相：码值锁存回放，仅复位沿出 [-] / fault, exit only on reset [-]
        ; // 锁存回放（R28） [-] / replay the latch only [-]
ELSE
    _iErr := 405; _eState := E_DL_TabCompState.eFault; // 非法相位兜底 [-] / illegal phase fallback [-]
END_CASE

// 段 3｜出口映射（名实双出口，同源赋值）
eState := _eState; // 状态出口 [-] / state outlet [-]
iErrCode := _iErr; // 故障码出口（锁存值） [-] / error code outlet [-]
iRejectCnt := _iRej; // 剔废计数出口 [片] / reject counter outlet [tablets]
xDone := xDoneInt AND NOT xDonePrev; // 完成单拍（内部锁存 → 出口映射） [-] / done one-shot [-]
xDonePrev := xDoneInt; // 本拍快照供下拍比较 [-] / snapshot for the next scan [-]
END_FUNCTION_BLOCK

(* ---- FB_DL_TabletWeightAutoCtl.st ---- *)
(*
  DL Factory R84 | FB_DL_TabletWeightAutoCtl
  功能：压片机片重自动控制：固定二十点滚动窗统计片重均值与标准差，按速度式 PI 出充填深度增量（死区＋限幅），单片按三倍标准差与上下公差判剔除，连续五片超差停机上报警。
  开源溯源：无（clean-room 自研，依据公开工艺公式与安全设计惯例，来源=行业通用公式+工程实践，许可证=MIT，借鉴点=公式结构与联锁分层）
  规则：R1-R16 全遵守
  ------------------------------------------------------------------
  分类 DL_Process ｜ 复杂度 cx4 ｜ 版本 v1.0.0 ｜ 平台 纯 IEC 61131-3（R_TRIG、LREAL、ENUM、CASE）
  边界一：只出充填深度指令与剔废脉冲，不驱动加料伺服、不控冲头行程、不执行剔废气缸（属主边界，执行由下层 PRG 完成）。
  边界二：滚动窗为定长二十槽环形缓冲（R15 显式定长），入窗与取窗同一存储；统计采用两遍法（先均值再离差平方和），
          分母为常量 20 与 19，结构性零除不可能；标准差取样本口径（分母 n−1）。
  边界三：判据次序为「先判后入窗」——单片离群判据使用入窗前的均值与标准差，避免本片自掩蔽把离群点拉回带内；
          剔除判定后该片仍入窗（工艺上已成型，属真实产出），故窗统计含被剔片，此口径写死在段 4 至段 6 顺序中。
  边界四：离群判据的三倍标准差门限仅在标准差大于零闸门限时生效；标准差为零（窗内全同）时只用公差判据，
          防「零标准差 → 任意微小偏差皆判离群」的假剔废群。
  边界五：调节量为速度式 PI 增量（du ＝ Kp·Δe ＋ Ki·e），积分效应内置于增量式，无独立积分累加器，
          故不存在积分饱和；累计指令的硬域钳定即为抗饱和的最终保障。死区为目标片重的 0.01 倍，死区内 e 取零，
          但 Δe 仍按零参与，使过零后不产生阶跃踢动。
  边界六：无效拍语义——目标片重不大于零、深度上下限越域、冲头压力低于下限、或任一浮点入参非有限 → xValid 出假、
          相位保持、调节量不出（深度指令保持上一值）；此三态均为信息级，故障级语义由 xStop 锁存位承担。
  量纲自检：片重 [mg]＝fWeightMg、fTargetMg、fTolUpMg、fTolDnMg、fMeanMg、fStdMg 同量纲；
          充填深度 [mm]＝fFillDepthMm、fDepthCmd、fDu、上下限；增益 Kp 单位 [mm/mg]、Ki 单位 [mm/mg]；
          压力 [kN]＝fForceKn 与 fForceMinKn。
  码表：本件全部码位为信息级（2801 目标片重越域、2802 深度限越域、2803 入参非有限、2804 压力低于下限、
        2805 连续超差停机、2806 非法相位）；信息级码每拍重算且不置 bError；停机锁存由 xStop 表达，故本件无 bError 出口（R187）。
  输出契约：fDepthCmd 为累计充填深度指令 [mm]（域内恒等于上下限之间）；xReject 为单拍剔除脉冲（统一出口映射）；
          xReady 在窗未满时为假且 fMeanMg 出 0（不出调节量）；iRejectCnt 为累计剔除片数 [片]，复位沿清零。
  修订记录：2026-11-24 v1.0.0 R84 首版（批 R84 · 序号 43）
*)

TYPE E_DL_TabWtState :
(
    eIdle     := 0, // 空闲：等使能与首片 / idle, waiting for the enable and the first tablet
    eSampling := 10, // 取样：窗未满，只统计不调节 / sampling, the window is filling and nothing is adjusted
    eAdjust   := 20, // 调节：窗已满，逐片出充填深度增量 / adjusting, the window is full and the depth is trimmed
    eReject   := 30, // 剔除：单拍过渡态，出剔除脉冲 / reject, a one scan transition emitting the reject pulse
    eStop     := 40  // 停机：连续超差锁存，复位沿解除 / stop, latched on consecutive deviations and cleared by the reset edge
);
END_TYPE

TYPE E_DL_TabWtCause :
(
    eNone      := 0, // 无成因 / no cause
    eTargetBad := 1, // 目标片重越域（信息级 2801）/ the target weight is out of domain, info grade 2801
    eLimitBad  := 2, // 充填深度上下限越域（信息级 2802）/ the depth limits are out of domain, info grade 2802
    eNotFinite := 3, // 入参非有限（信息级 2803）/ a non-finite input, info grade 2803
    eForceLow  := 4, // 冲头压力低于下限（信息级 2804）/ the punch force is below its floor, info grade 2804
    eConsBad   := 5, // 连续超差停机（信息级 2805）/ consecutive deviations tripped the machine, info grade 2805
    ePhaseBad  := 6  // 非法相位（信息级 2806）/ an illegal phase, info grade 2806
);
END_TYPE

FUNCTION_BLOCK FB_DL_TabletWeightAutoCtl
VAR CONSTANT
    DL_TWC_WIN         : INT := 20;       // 滚动窗点数 [点] / the rolling window length [point]
    DL_TWC_WIN_CAP     : INT := 20;       // 缓冲槽数（下标 0..19，与窗点数一致）[槽] / the buffer slots, subscripts 0..19 [slot]
    DL_TWC_DEN_N       : LREAL := 20.0;   // 均值分母（常量，结构性非零）[-] / the mean denominator as a constant [-]
    DL_TWC_DEN_N1      : LREAL := 19.0;   // 样本方差分母 n−1（常量）[-] / the sample variance denominator [-]
    DL_TWC_KP          : LREAL := 0.020;  // 比例增益 [mm/mg] / the proportional gain [mm/mg]
    DL_TWC_KI          : LREAL := 0.004;  // 积分增益（速度式内的积分项）[mm/mg] / the integral gain inside the velocity form [mm/mg]
    DL_TWC_DEADBAND_FRAC : LREAL := 0.01; // 死区带宽（目标片重的倍数）[-] / the dead band as a fraction of the target [-]
    DL_TWC_STEP_MM     : LREAL := 0.05;   // 单次调节限幅 [mm] / the per shot adjustment step limit [mm]
    DL_TWC_SIGMA_K     : LREAL := 3.0;    // 离群判据的标准差倍数 [-] / the sigma multiplier of the outlier test [-]
    DL_TWC_CONS_MAX    : INT := 5;        // 连续超差停机点数 [片] / the consecutive deviation trip count [tablet]
    DL_TWC_EPS         : LREAL := 1.0E-9; // 零闸与零判定门限 [-] / the zero guard and zero test threshold [-]
END_VAR
VAR_INPUT
    bEnable       : BOOL := TRUE;    // 使能，失能回空闲且不再调节 [-] / enable, a disable returns to idle and stops trimming
    bReset        : BOOL := FALSE;   // 复位上升沿清停机锁存与全部计数 [-] / reset rising edge clears the stop latch and the counters
    bPieceValid   : BOOL := FALSE;   // 新片有效（脉冲或电平，取上升沿）[-] / a valid tablet, its rising edge is consumed
    fWeightMg     : LREAL := 500.0;  // 实测片重 [mg] / the measured tablet weight [mg]
    fTargetMg     : LREAL := 500.0;  // 目标片重 [mg] / the target tablet weight [mg]
    fTolUpMg      : LREAL := 10.0;   // 上公差 [mg] / the upper tolerance [mg]
    fTolDnMg      : LREAL := 10.0;   // 下公差 [mg] / the lower tolerance [mg]
    fFillDepthMm  : LREAL := 8.00;   // 充填深度反馈 [mm] / the fill depth feedback [mm]
    fFillDepthMinMm : LREAL := 4.00; // 充填深度下限 [mm] / the fill depth lower limit [mm]
    fFillDepthMaxMm : LREAL := 14.0; // 充填深度上限 [mm] / the fill depth upper limit [mm]
    fForceKn      : LREAL := 30.0;   // 冲头压力 [kN] / the punch force [kN]
    fForceMinKn   : LREAL := 5.00;   // 冲头压力下限（低于即无效拍）[kN] / the punch force floor [kN]
END_VAR
VAR_OUTPUT
    fDepthCmd    : LREAL := 0.0;  // 充填深度指令（累计）[mm] / the fill depth command, accumulated [mm]
    fMeanMg      : LREAL := 0.0;  // 窗内片重均值（窗未满出 0）[mg] / the window mean, zero until the window is full [mg]
    fStdMg       : LREAL := 0.0;  // 窗内片重样本标准差 [mg] / the window sample standard deviation [mg]
    fDevMg       : LREAL := 0.0;  // 本片相对上拍均值的偏差 [mg] / the deviation of the tablet against the previous mean [mg]
    iRejectCnt   : DINT := 0;     // 累计剔除片数 [片] / the accumulated reject count [tablet]
    nWinFill     : INT := 0;      // 窗内已填点数 [点] / the filled window points [point]
    xReject      : BOOL := FALSE; // 单拍剔除脉冲（统一出口映射）[-] / the one scan reject pulse
    xStop        : BOOL := FALSE; // 停机锁存（连续超差，复位沿清除）[-] / the stop latch cleared by the reset edge
    xReady       : BOOL := FALSE; // 窗已满且可出调节量 [-] / the window is full and a trim may be issued
    eState       : E_DL_TabWtState := E_DL_TabWtState.eIdle; // 相位出口 [枚举] / the phase outlet [enum]
    iErrCode     : INT := 0;      // 信息级码（每拍重算，非锁存）[码] / the info grade code, recomputed every scan [code]
    xValid       : BOOL := FALSE; // 本拍输入可信 [-] / the inputs of this scan are trustworthy
END_VAR
VAR
    rtPiece    : R_TRIG; // 新片沿实例（无量纲）[-] / the tablet edge refreshed unconditionally
    rtReset    : R_TRIG; // 复位沿实例（无量纲）[-] / the reset edge refreshed unconditionally
    _eState    : E_DL_TabWtState := E_DL_TabWtState.eIdle; // 内部相位（枚举，无量纲）[-] / the internal phase, the only CASE target
    _aBuf      : ARRAY[0..19] OF LREAL; // 片重环形缓冲（定长二十槽，R15）[mg] / the ring buffer of the weights [mg]
    _iHead     : INT := 0;    // 下一点写入槽号（0..19）[槽] / the next write slot [slot]
    _iFill     : INT := 0;    // 已填点数（封顶二十）[点] / the filled points capped at twenty [point]
    _i         : INT := 0;    // 遍历下标 [-] / the traversal index
    _iConsBad  : INT := 0;    // 连续超差片数 [片] / the consecutive deviating count [tablet]
    _iErrTmp   : INT := 0;    // 本拍信息级码暂存 [码] / the scan info code scratch [code]
    _iRejAcc   : DINT := 0;   // 剔除计数累加（唯一写入点）[片] / the reject accumulator, the only write point [tablet]
    _bInit     : BOOL := FALSE; // 首扫初始化完成标志（R310）[-] / the first scan initialisation flag
    _bFinOk    : BOOL := FALSE; // 全部浮点入参有限 [-] / every floating input is finite
    _bTgtOk    : BOOL := FALSE; // 目标片重与公差域内 [-] / the target and the tolerances are inside the domain
    _bLimOk    : BOOL := FALSE; // 深度上下限域内 [-] / the depth limits are inside the domain
    _bForceOk  : BOOL := FALSE; // 冲头压力不低于下限 [-] / the punch force is at or above its floor
    _bWinFull  : BOOL := FALSE; // 窗已填满（可统计可调节）[-] / the window is full
    _bReject   : BOOL := FALSE; // 本片剔除判据结果 [-] / the reject verdict of the tablet
    _bOverTol  : BOOL := FALSE; // 本片超公差（参与连续计数）[-] / the tablet broke the tolerance
    _bRejOut   : BOOL := FALSE; // 单拍剔除位（段 0 预清，出口映射）[-] / the one scan reject bit
    _bStopLch  : BOOL := FALSE; // 停机锁存位（唯一清除：复位沿）[-] / the stop latch cleared by the reset edge only
    _bAdjOk    : BOOL := FALSE; // 本拍允许调节（状态量与窗满合取）[-] / the trim permit from the state and the window
    _fSum      : LREAL := 0.0;  // 窗内片重和 [mg] / the window sum [mg]
    _fMean     : LREAL := 0.0;  // 窗内均值（本拍计算）[mg] / the window mean of this scan [mg]
    _fDev      : LREAL := 0.0;  // 单点离差（窗统计遍历用）[mg] / the single point deviation used by the traversal [mg]
    _fDevPiece : LREAL := 0.0;  // 本片相对上拍均值的偏差（判据与诊断）[mg] / the tablet deviation against the previous mean [mg]
    _fVar      : LREAL := 0.0;  // 窗内样本方差 [mg²] / the window sample variance [mg^2]
    _fStd      : LREAL := 0.0;  // 窗内样本标准差 [mg] / the window sample standard deviation [mg]
    _fMeanPrev : LREAL := 0.0;  // 上拍均值快照（判据用，不含本片）[mg] / the previous mean snapshot used by the verdict [mg]
    _fStdPrev  : LREAL := 0.0;  // 上拍标准差快照（判据用）[mg] / the previous deviation snapshot used by the verdict [mg]
    _fErr      : LREAL := 0.0;  // 片重偏差（目标减均值，正为偏轻）[mg] / the weight error, positive means too light [mg]
    _fErrEff   : LREAL := 0.0;  // 死区处理后的偏差 [mg] / the error after the dead band [mg]
    _fErrPrev  : LREAL := 0.0;  // 上次调节的偏差快照 [mg] / the error snapshot of the last trim [mg]
    _fBand     : LREAL := 0.0;  // 死区带宽 [mg] / the dead band width [mg]
    _fDu       : LREAL := 0.0;  // 速度式 PI 增量（限幅前）[mm] / the velocity form increment before limiting [mm]
    _fCmd      : LREAL := 0.0;  // 充填深度指令累加（唯一写入点）[mm] / the depth command accumulator [mm]
END_VAR
// 段 0｜出口预置：全部出口先赋安全侧值，任何路径不留未初始化输出
xValid := FALSE; // 有效性预置假 / validity preset false
xReady := _bWinFull AND bEnable; // 就绪位预置（窗满且使能）/ the ready bit preset
xReject := FALSE; // 剔除脉冲预置假（本拍重新判定）/ the reject pulse preset false
xStop := _bStopLch; // 停机锁存回放 / replay the stop latch
fDepthCmd := _fCmd; // 深度指令回放上一值（无效拍保持）/ replay the last depth command
fMeanMg := 0.0; // 均值预置零（窗未满契约）/ the mean preset zero
fStdMg := 0.0; // 标准差预置零 / the standard deviation preset zero
fDevMg := 0.0; // 偏差预置零 / the deviation preset zero
iRejectCnt := _iRejAcc; // 剔除计数回放 / replay the reject count
nWinFill := _iFill; // 窗内点数回放 / replay the filled points
eState := _eState; // 相位回放 / replay the phase
iErrCode := 0; // 信息级码预置零（本拍重算）/ the info code preset zero
_bRejOut := FALSE; // 单拍剔除位预清零（FB32-1：仅单拍标志可预清）/ preclear the one scan reject bit
_bReject := FALSE; // 单拍剔除判据预清 / preclear the reject verdict
_bOverTol := FALSE; // 单拍超公差判据预清 / preclear the tolerance verdict
_iErrTmp := 0; // 单拍码暂存预清 / preclear the code scratch
// 段 1｜非有限闸：NaN 自反比较、Inf 差值自减双判，逐项枚举八个浮点入参（R79、R272）
_bFinOk := (fWeightMg = fWeightMg) AND ((fWeightMg - fWeightMg) = (fWeightMg - fWeightMg)) // 片重有限 [-] / the weight is finite
    AND (fTargetMg = fTargetMg) AND ((fTargetMg - fTargetMg) = (fTargetMg - fTargetMg)) // 目标片重有限 [-] / the target is finite
    AND (fTolUpMg = fTolUpMg) AND ((fTolUpMg - fTolUpMg) = (fTolUpMg - fTolUpMg)) // 上公差有限 [-] / the upper tolerance is finite
    AND (fTolDnMg = fTolDnMg) AND ((fTolDnMg - fTolDnMg) = (fTolDnMg - fTolDnMg)) // 下公差有限 [-] / the lower tolerance is finite
    AND (fFillDepthMm = fFillDepthMm) AND ((fFillDepthMm - fFillDepthMm) = (fFillDepthMm - fFillDepthMm)) // 深度反馈有限 [-] / the depth feedback is finite
    AND (fFillDepthMinMm = fFillDepthMinMm) AND ((fFillDepthMinMm - fFillDepthMinMm) = (fFillDepthMinMm - fFillDepthMinMm)) // 深度下限有限 [-] / the depth floor is finite
    AND (fFillDepthMaxMm = fFillDepthMaxMm) AND ((fFillDepthMaxMm - fFillDepthMaxMm) = (fFillDepthMaxMm - fFillDepthMaxMm)) // 深度上限有限 [-] / the depth ceiling is finite
    AND (fForceKn = fForceKn) AND ((fForceKn - fForceKn) = (fForceKn - fForceKn)) // 冲头压力有限 [-] / the punch force is finite
    AND (fForceMinKn = fForceMinKn) AND ((fForceMinKn - fForceMinKn) = (fForceMinKn - fForceMinKn)); // 压力下限有限 [-] / the force floor is finite
// 段 2｜组态域闸：目标片重正定、公差非负、深度上限大于下限、压力下限非负（R151、FB51-2）
_bTgtOk := (fTargetMg > 0.0) AND (fTolUpMg >= 0.0) AND (fTolDnMg >= 0.0); // 目标与公差域闸 [-] / the target and the tolerance gates
_bLimOk := (fFillDepthMinMm > 0.0) AND (fFillDepthMaxMm > fFillDepthMinMm); // 深度域闸（上限严格大于下限）[-] / the depth domain gate
_bForceOk := (fForceMinKn >= 0.0) AND (fForceKn >= fForceMinKn); // 压力域闸 [-] / the force domain gate
IF NOT _bFinOk THEN _iErrTmp := 2803; // 信息级：入参非有限 / the info code for a non-finite input
ELSIF NOT _bTgtOk THEN _iErrTmp := 2801; // 信息级：目标片重越域 / the info code for a bad target
ELSIF NOT _bLimOk THEN _iErrTmp := 2802; // 信息级：深度限越域 / the info code for bad depth limits
ELSIF NOT _bForceOk THEN _iErrTmp := 2804; // 信息级：压力低于下限 / the info code for a low punch force
END_IF
// 段 3｜沿检测无条件周期刷新（R7）
rtPiece(CLK := bPieceValid); // 新片沿无条件刷新 / unconditional refresh of the tablet edge
rtReset(CLK := bReset); // 复位沿无条件刷新 / unconditional refresh of the reset edge
// 段 4｜首扫初始化与复位沿同块，作用域逐项声明（R310、R311）
IF (NOT _bInit) OR rtReset.Q THEN // 首扫一拍或复位沿 / the first scan or the reset edge
    _bInit := TRUE; // 首扫完成标志 / the first scan flag
    _bStopLch := FALSE; // 作用域一：清停机锁存（唯一清除边，R188）/ scope one, clear the stop latch
    _iRejAcc := 0; _iConsBad := 0; // 作用域二：清剔除计数与连续超差计数 / scope two, clear the counters
    _iHead := 0; _iFill := 0; // 作用域二：缓冲复位 / scope two, reset the buffer
    _fMeanPrev := 0.0; _fStdPrev := 0.0; _fErrPrev := 0.0; // 作用域三：清统计与调节快照 / scope three, clear the snapshots
    _fCmd := fFillDepthMm; // 作用域三：指令基准取当前反馈 [mm] / scope three, the command base is the feedback [mm]
    IF _fCmd < fFillDepthMinMm THEN _fCmd := fFillDepthMinMm; END_IF // 基准下限钳定 / clamp the base low
    IF _fCmd > fFillDepthMaxMm THEN _fCmd := fFillDepthMaxMm; END_IF // 基准上限钳定 / clamp the base high
    _eState := E_DL_TabWtState.eIdle; // 作用域二：迁回空闲相 / scope two, migrate to idle
END_IF
// 段 5｜单片剔除判据：先用上拍统计（不含本片），3σ 门限仅在标准差有效时生效（边界四）
IF rtPiece.Q AND _bFinOk AND _bTgtOk THEN // 新片且目标与入参可信 / a new tablet with a trustworthy target
    _fDevPiece := fWeightMg - _fMeanPrev; // 本片偏差 [mg] / the deviation of the tablet [mg]
    IF _fStdPrev > DL_TWC_EPS THEN // 标准差有效才用三倍标准差判据 / the sigma test only with a valid deviation
        IF ABS(_fDevPiece) > (DL_TWC_SIGMA_K * _fStdPrev) THEN _bReject := TRUE; END_IF // 三倍标准差离群 / the three sigma outlier
    END_IF
    IF fWeightMg > (fTargetMg + fTolUpMg) THEN _bReject := TRUE; _bOverTol := TRUE; END_IF // 上公差越限（方向分列）/ the upper tolerance breach
    IF fWeightMg < (fTargetMg - fTolDnMg) THEN _bReject := TRUE; _bOverTol := TRUE; END_IF // 下公差越限（方向分列）/ the lower tolerance breach
    IF _bReject THEN // 判为剔除 / judged as a reject
        _iRejAcc := _iRejAcc + 1; // 累计剔除片数（唯一写入点）/ the only write point of the reject count
        _bRejOut := TRUE; // 置单拍剔除位（出口统一映射，R187）/ raise the one scan reject bit
    END_IF
    IF _bOverTol THEN _iConsBad := _iConsBad + 1; ELSE _iConsBad := 0; END_IF // 连续超差净额计数（单点写入）/ the net consecutive count
    IF _iConsBad >= DL_TWC_CONS_MAX THEN _bStopLch := TRUE; END_IF // 连续五片超差：锁存停机 / five in a row latch the stop
END_IF
// 段 6｜入窗：环形推进（禁 MOD，R140 委托边界），写入值已过有限闸
IF rtPiece.Q AND _bFinOk THEN // 新片且入参可信 / a new tablet with trustworthy inputs
    IF (_iHead >= 0) AND (_iHead <= (DL_TWC_WIN_CAP - 1)) THEN // 写槽下标先夹取（R4 越界防御）/ clamp the slot subscript first
        _aBuf[_iHead] := fWeightMg; // 写当前槽 [mg] / write the current slot [mg]
    END_IF
    IF _iHead >= (DL_TWC_WIN_CAP - 1) THEN _iHead := 0; ELSE _iHead := _iHead + 1; END_IF // 环形推进 / advance the ring
    IF _iFill < DL_TWC_WIN_CAP THEN _iFill := _iFill + 1; END_IF // 已填点数封顶 / cap the filled points
END_IF
_bWinFull := _iFill >= DL_TWC_WIN; // 窗满判据 / the window full verdict
// 段 7｜窗统计：两遍法（均值 → 离差平方和），分母为常量 20 与 19（结构性零除不可能）
IF _bWinFull THEN // 窗满才统计 / statistics only with a full window
    _fSum := 0.0; // 求和累加清零 / clear the sum
    FOR _i := 0 TO (DL_TWC_WIN_CAP - 1) DO // 第一遍：求和（定长字面界）/ pass one, the sum
        _fSum := _fSum + _aBuf[_i]; // 逐槽累加 [mg] / accumulate slot by slot [mg]
    END_FOR
    _fMean := _fSum / DL_TWC_DEN_N; // 均值 [mg] / the mean [mg]
    _fVar := 0.0; // 离差平方和清零 / clear the squared deviations
    FOR _i := 0 TO (DL_TWC_WIN_CAP - 1) DO // 第二遍：离差平方和（定长字面界）/ pass two, the squared deviations
        _fDev := _aBuf[_i] - _fMean; // 单点离差 [mg] / the single point deviation [mg]
        _fVar := _fVar + (_fDev * _fDev); // 累加平方 [mg²] / accumulate the square [mg^2]
    END_FOR
    _fVar := _fVar / DL_TWC_DEN_N1; // 样本方差 [mg²] / the sample variance [mg^2]
    IF _fVar < 0.0 THEN _fVar := 0.0; END_IF // 舍入残差负方差钳零 / clamp the rounding residual
    _fStd := SQRT(_fVar); // 样本标准差 [mg] / the sample standard deviation [mg]
    IF NOT (_fStd = _fStd) THEN _fStd := 0.0; END_IF // 标准差 NaN 兜底 / the NaN fallback
    IF (_fStd - _fStd) <> (_fStd - _fStd) THEN _fStd := 0.0; END_IF // 标准差 Inf 兜底 / the Inf fallback
    _fMeanPrev := _fMean; // 均值快照供下一片判据（不含下一片）/ the mean snapshot for the next verdict
    _fStdPrev := _fStd; // 标准差快照供下一片判据 / the deviation snapshot for the next verdict
END_IF
// 段 8｜速度式 PI 调节：窗满、新片、使能、未锁存、输入可信五条件齐备才出增量（状态量门控，R99）
_bAdjOk := _bWinFull AND bEnable AND (NOT _bStopLch) AND _bFinOk AND _bTgtOk; // 调节许可合取 / the trim permit
IF _bAdjOk AND rtPiece.Q THEN // 仅在窗满后的每片调节一次 / trim once per tablet after the window filled
    _fErr := fTargetMg - _fMean; // 片重偏差 [mg]，正为偏轻需加深 / the error, positive means too light
    _fBand := fTargetMg * DL_TWC_DEADBAND_FRAC; // 死区带宽 [mg] / the dead band width [mg]
    IF ABS(_fErr) <= _fBand THEN _fErrEff := 0.0; ELSE _fErrEff := _fErr; END_IF // 死区内偏差取零 / zero the error inside the dead band
    _fDu := (DL_TWC_KP * (_fErrEff - _fErrPrev)) + (DL_TWC_KI * _fErrEff); // 速度式 PI 增量 [mm] / the velocity form increment [mm]
    IF _fDu > DL_TWC_STEP_MM THEN _fDu := DL_TWC_STEP_MM; ELSIF _fDu < (0.0 - DL_TWC_STEP_MM) THEN _fDu := (0.0 - DL_TWC_STEP_MM); END_IF // 单次调节双向限幅 / the two sided step limit
    IF NOT (_fDu = _fDu) THEN _fDu := 0.0; END_IF // 增量 NaN 兜底（拒收不外抛）/ the NaN fallback
    IF (_fDu - _fDu) <> (_fDu - _fDu) THEN _fDu := 0.0; END_IF // 增量 Inf 兜底 / the Inf fallback
    _fCmd := _fCmd + _fDu; // 累计指令（唯一写入点）[mm] / the only write point of the command [mm]
    IF _fCmd > fFillDepthMaxMm THEN _fCmd := fFillDepthMaxMm; END_IF // 上限硬钳（抗饱和终保）/ the hard clamp high
    IF _fCmd < fFillDepthMinMm THEN _fCmd := fFillDepthMinMm; END_IF // 下限硬钳 / the hard clamp low
    _fErrPrev := _fErrEff; // 偏差快照（供下一次差分）/ the error snapshot for the next difference
END_IF
// 段 9｜相位状态机：ENUM ＋ CASE ＋ ELSE 非法相位兜底（R6、R128）
CASE _eState OF
E_DL_TabWtState.eIdle: // 空闲相：退出条件三（使能丢失驻留、锁存升停机、首片进取样）
    IF _bStopLch THEN // 停机锁存已置 / the stop latch is set
        _eState := E_DL_TabWtState.eStop; // 迁停机相 / migrate to stop
    ELSIF bEnable AND rtPiece.Q THEN // 使能且首片到达 / enabled with the first tablet
        _eState := E_DL_TabWtState.eSampling; // 迁取样相 / migrate to sampling
    END_IF
E_DL_TabWtState.eSampling: // 取样相：退出条件四（失能、锁存、剔除、窗满）
    IF NOT bEnable THEN // 使能丢失 / the enable was lost
        _eState := E_DL_TabWtState.eIdle; // 回空闲 / back to idle
    ELSIF _bStopLch THEN // 停机锁存已置 / the stop latch is set
        _eState := E_DL_TabWtState.eStop; // 迁停机相 / migrate to stop
    ELSIF _bRejOut THEN // 本片判剔除（拍 N 进入：本片判据命中；本拍行为：拒收并出脉冲；拍 N+1 转出：回取样或调节）
        _eState := E_DL_TabWtState.eReject; // 迁剔除过渡相 / migrate to the reject transition
    ELSIF _bWinFull THEN // 窗已满（本拍不调节，下一片起调节）/ the window is full
        _eState := E_DL_TabWtState.eAdjust; // 迁调节相 / migrate to adjusting
    END_IF
E_DL_TabWtState.eAdjust: // 调节相：退出条件三（失能、锁存、剔除）
    IF NOT bEnable THEN // 使能丢失 / the enable was lost
        _eState := E_DL_TabWtState.eIdle; // 回空闲 / back to idle
    ELSIF _bStopLch THEN // 停机锁存已置 / the stop latch is set
        _eState := E_DL_TabWtState.eStop; // 迁停机相 / migrate to stop
    ELSIF _bRejOut THEN // 本片判剔除 / the tablet is a reject
        _eState := E_DL_TabWtState.eReject; // 迁剔除过渡相 / migrate to the reject transition
    END_IF
E_DL_TabWtState.eReject: // 剔除过渡相：本拍不出调节量，只等本拍之后转出
    IF _bStopLch THEN // 停机锁存已置 / the stop latch is set
        _eState := E_DL_TabWtState.eStop; // 迁停机相 / migrate to stop
    ELSIF _bWinFull THEN // 窗已满：回调节相 / the window is full, back to adjusting
        _eState := E_DL_TabWtState.eAdjust; // 回调节相 / back to adjusting
    ELSE // 窗未满：回取样相 / the window is not full, back to sampling
        _eState := E_DL_TabWtState.eSampling; // 回取样相 / back to sampling
    END_IF
E_DL_TabWtState.eStop: // 停机相：锁存驻留，唯一解除为复位沿（段 4 已迁回空闲）
    IF NOT _bStopLch THEN // 锁存已被复位沿清除 / the latch was cleared by the reset edge
        _eState := E_DL_TabWtState.eIdle; // 回空闲 / back to idle
    END_IF
ELSE // 非法相位兜底（R6、R128）
    _eState := E_DL_TabWtState.eStop; // 落停机安全相 / fall back to the safe stop phase
    _iErrTmp := 2806; // 信息级非法相位码 / the info grade illegal phase code
END_CASE
// 段 10｜统一出口：单点映射，剔除脉冲与停机位同源派生（R191、FB51-8）
eState := _eState; // 相位单点映射 / the single point mapping of the phase
xReject := _bRejOut; // 剔除脉冲单点映射（单拍，段 0 已预清）/ the one scan reject pulse
xStop := _bStopLch; // 停机锁存单点映射 / the single point mapping of the stop latch
fDepthCmd := _fCmd; // 深度指令单点映射 [mm] / the single point mapping of the depth command [mm]
nWinFill := _iFill; // 窗内点数单点映射 / the single point mapping of the filled points
iRejectCnt := _iRejAcc; // 剔除计数单点映射 / the single point mapping of the reject count
IF _bWinFull THEN // 窗满才外抛统计量 / publish the statistics only with a full window
    fMeanMg := _fMean; // 均值 [mg] / the mean [mg]
    fStdMg := _fStd; // 标准差 [mg] / the standard deviation [mg]
ELSE // 窗未满：按契约出零（不出调节量）/ not full, the contract demands zeros
    fMeanMg := 0.0; // 均值出零 / the mean goes to zero
    fStdMg := 0.0; // 标准差出零 / the deviation goes to zero
END_IF
fDevMg := _fDevPiece; // 本片偏差（诊断用）[mg] / the tablet deviation for diagnostics [mg]
xReady := _bWinFull AND bEnable AND (NOT _bStopLch); // 就绪位：窗满、使能、未锁存 / the ready bit
IF _bStopLch AND (_iErrTmp = 0) THEN _iErrTmp := 2805; END_IF // 停机原因码（信息级，锁存语义由 xStop 承担）/ the stop cause code
iErrCode := _iErrTmp; // 信息级码单点映射（每拍重算，不锁存）/ the info code mapping
xValid := _bFinOk AND _bTgtOk AND _bLimOk AND _bForceOk AND (_iErrTmp = 0); // 有效性：四闸通过且无信息级码
END_FUNCTION_BLOCK

(* ---- FB_DL_TaktPaceMonitor.st ---- *)
(*
  ==================================================================
  组件名 Component  : FB_DL_TaktPaceMonitor
  分类   Category   : DL_Process
  前缀   Naming     : FB_DL_ ｜ b/n/u/f/t/e 类型前缀制（R265）
  版本   Version    : 1.0.2
  功能   Purpose    : 节拍 / 进度落后监视（ISO 22400-2 公开口径）：bCycleDone
                      两脉冲间隔测实际节拍，EWMA（系数 fAlpha ∈ (0,1]）平滑
                      为 fTaktActS；fPaceDevPct = (实际 − 目标)/目标 × 100，
                      正值即落后（bBehind）。tEvalWindow 评估窗滚动统计窗内
                      产量对目标产量的缺口 uQtyBacklog（溢出钳位 + 信息码）。
                      首件前不出数（bValid=FALSE）；窗内零产出是合法观测——
                      缺口 = 窗内目标产量全额（分母侧显式判，不除以产量）。
  来源   Source     : self-std（ISO 22400-2 节拍/缺口公开口径，零源码复制，
                      术语与公式口径为公开标准条款）
  互引   Cross-ref  : FB_DL_CycleTimeMeasure（同族周期测量件：其 uCycleLast
                      可作本件目标节拍整定参考）；FB_DL_OeeCalculator
                      （下游 KPI 件：本件 fPaceDevPct / uQtyBacklog 可作其
                      性能类输入）
  平台   Platform   : 纯 IEC 61131-3（R_TRIG/LREAL 四则/TIME 比较与整转）
  依赖   Depends    : 仅 Standard.library（R_TRIG 属标准件）；TIME_TO_DINT
                      属 IEC 标准类型转换
  设计偏差 Deviation: 时间基准按本库「时间注入」纪律：新增输入 fCallCycleS
                      （调用方注入扫描周期 [s]，FB_DL_CycleTimeMeasure 语义），
                      本件不读平台时刻函数；tEvalWindow 以 TIME_TO_DINT 转
                      毫秒参与闸与滚动判据（TIME 本义即 ms，三平台一致）。
  红线   Redline    : R1 零全局/VAR_EXTERNAL/R2 零 %I/%Q/R3 纯 IEC 标准
                      R4 分母三闸（目标节拍 / 目标+实际差 / 窗长）显式判 +
                      溢出钳位显式 + 非有限闸 + 输出域显式
                      R5 全变量双语同行注释/R6 配置故障为电平面无状态机
                      （CASE 不适用，头注说明）/R7 rtCycle 段 0 无条件刷新
                      R8 容差与阈值常量化
  契约   Contract   : 配置故障（码 01/02）为电平面（当拍复判，非锁存）：故障
                      拍 bValid=FALSE、输出全部冻结保持、bError=TRUE；恢复
                      即恢复。失能相（bEnable=FALSE）串清账：窗内累计清零、
                      上一脉冲基准撤销、bValid=FALSE（R 失能清账条款）。
  错误码 Codes      : 01【故障级】目标节拍配置非法（≤ 0 或非有限）、评估窗
                      非法（≤ T#0MS）或扫描周期注入非法（≤ 0 / 非有限，
                      v1.0.1 将窗面/计时面并入本码，修静默降级）
                      02【故障级】平滑系数 fAlpha 域外（须 (0,1]）或非有限
                      03【信息级】缺口/窗内计数溢出钳位（饱和于 UDINT 上限）
  码位反证 Note     : 01/02 分立依据（R90）：01 在目标面与窗面、02 在平滑
                      系数面可观测，整定入口不同；03 为信息级不置 bError，
                      与 01/02 双通道可区分；窗长非法并入 01 的反证：窗长
                      与目标同为「节拍推进判据」的标定面，处置同形（冻结
                      + 拒推进），输出组合不可区分。
  验收   Acceptance : V1 稳定 60s 节拍 → fTaktActS→60，fPaceDevPct 随目标
                      ｜ V2 目标 50s 实际 60s → bBehind=TRUE ｜ V3 alpha=0
                      或 1.5 → 码 02 ｜ V4 首件前 bValid=FALSE ｜ V5 窗内
                      零产出 → 缺口 = 窗内目标产量（码面无 03）｜ V6 超长窗
                      小目标 → 缺口钳上限 + 码 03 ｜ V7 失能 → 全清账
  变更   Revision   : 2026-11-22  v1.0.0  R66 首版（编码阶段批 4 序 10）
                      2026-11-22  v1.0.1  R66 终审就地修（1 中）：窗面/计时
                      基准面失效原走静默降级（bValid=FALSE 但不置 bError
                      不置码，R258 家族），并入码 01 电平面出口。
                      2026-11-22  v1.0.2  R67 点修（L4）：段 5 fExpectR 闸界
                      由 UDINT 域 4.294967295E9 前移至 DINT 中转域上界
                      2147483647（常量 TPM_DINT_MAX，与 TIME_TO_DINT /
                      LREAL_TO_DINT 转换链中转域 2^31−1 对齐，窗/目标比 >
                      2.1e9 s 组态下原转换链溢出可达）；M1 码 01 判式
                      （NOT _bTgtOk OR NOT _bTimeOk）维持 v1.0.1 不回退。
  ==================================================================
*)
FUNCTION_BLOCK FB_DL_TaktPaceMonitor
VAR_INPUT
    bCycleDone   : BOOL := FALSE;    // 完工脉冲输入（上升沿计件与测节拍）[-] / the cycle done pulse, counted on the rising edge
    fTaktTargetS : LREAL := 60.0;    // 目标节拍 [s]，须 > 0 且有限 / the takt target, positive and finite
    bEnable      : BOOL := FALSE;    // 使能，FALSE 失能清账（头注契约）[-] / the enable, false clears the books
    fAlpha       : LREAL := 0.2;     // EWMA 平滑系数 [-]，有效域 (0,1] / the EWMA factor, inside zero exclusive to one inclusive
    tEvalWindow  : TIME := T#60M;    // 评估窗长 [ms]（TIME 本义 ms），须 > 0 / the evaluation window length, must be positive
    fCallCycleS  : LREAL := 0.01;    // 调用方注入扫描周期 [s]，须 > 0 / the caller injected scan cycle in seconds
END_VAR
VAR_OUTPUT
    fTaktActS    : LREAL := 0.0;     // EWMA 实际节拍 [s]（首件前保持 0 并 bValid=FALSE）/ the EWMA actual takt [s]
    fPaceDevPct  : LREAL := 0.0;     // 进度偏差 [(实际−目标)/目标×100]，正=落后 [%] / the pace deviation percent, positive is behind
    uQtyBacklog  : UDINT := UDINT#0; // 窗口产量缺口 [件]（溢出钳位）/ the window production backlog, saturated
    bBehind      : BOOL := FALSE;    // 落后指示（fPaceDevPct > 0）[-] / the behind indicator
    bValid       : BOOL := FALSE;    // 输出有效标志（首件前=FALSE）[-] / the output validity, false before the first piece
    bError       : BOOL := FALSE;    // 配置故障标志（电平面，恢复即清，R45 配对）/ the configuration fault flag, per scan level
    uErrorId     : UDINT := 16#0000_0000; // 错误码，0=正常，01/02/03 见头注 [码] / the error code [code]
END_VAR
VAR
    rtCycle      : R_TRIG;           // 完工沿实例，段 0 无条件刷新 / the cycle edge instance refreshed unconditionally
    _bHasPrev    : BOOL := FALSE;    // 上一完工脉冲基准是否存在（首件判据）[-] / the previous pulse baseline flag
    _fSinceS     : LREAL := 0.0;     // 距上一完工脉冲的累计时长 [s] / the time since the previous pulse [s]
    _bTaktInit   : BOOL := FALSE;    // EWMA 是否已初始化（首个有效间隔直赋）[-] / the EWMA seeded flag
    _fWinAccMs   : LREAL := 0.0;     // 评估窗累计时长 [ms] / the window elapsed accumulator [ms]
    _uQtyWin     : UDINT := UDINT#0; // 窗内实际产量 [件] / the in window actual quantity [pc]
    _fWinLimMs   : LREAL := 0.0;     // 评估窗长整定 [ms]（TIME 转 LREAL 缓存）/ the window limit cached from TIME [ms]
    _bTgtOk      : BOOL := FALSE;    // 本拍目标有效性 [-] / the per scan target validity
    _bAlphaOk    : BOOL := FALSE;    // 本拍平滑系数有效性 [-] / the per scan alpha validity
    _bTimeOk     : BOOL := FALSE;    // 本拍计时基准有效性 [-] / the per scan time base validity
    _nExpect     : UDINT := UDINT#0; // 窗内目标产量工作寄存器 [件] / the in window expected quantity register
    _bQtySat     : BOOL := FALSE;    // 本拍溢出钳位信息位（单拍）/ the per scan saturation info bit
    fInterval    : LREAL := 0.0;     // 当前完工间隔工作寄存器 [s] / the current interval working register [s]
    fExpectR     : LREAL := 0.0;     // 窗内目标产量实数工作寄存器 [件] / the expected quantity as real [pc]
END_VAR
VAR CONSTANT
    TPM_FIN_MAX   : LREAL := 1.7976931348623157E308; // LREAL 有限上限 / the finite LREAL limit
    TPM_EPS       : LREAL := 1.0E-9;   // 到达与零判容差 [无量纲] / the tolerance for zero tests
    TPM_U_MAX     : UDINT := 4294967295; // UDINT 上限哨兵 [件] / the UDINT ceiling sentinel
    TPM_DINT_MAX  : LREAL := 2147483647.0; // DINT 中转域上界 2^31-1（实数钳界，v1.0.2 前移）/ the DINT transit domain ceiling
    TPM_ERR_NONE  : UDINT := 16#0000_0000; // 无错误 [码] / no error [code]
    TPM_ERR_TGT   : UDINT := 16#0000_0001; // 码 01：目标/窗配置非法 / code 01, target or window illegal
    TPM_ERR_ALPHA : UDINT := 16#0000_0002; // 码 02：平滑系数域外 / code 02, alpha out of domain
    TPM_ERR_SAT   : UDINT := 16#0000_0003; // 码 03：缺口/计数溢出钳位（信息级）/ code 03, saturation, info level
END_VAR

(*------------------------------------------------------------------------------
 * 段 0｜沿检测无条件刷新区（红线 R7）：严禁移入 IF / CASE
 *      The edge instance refreshes unconditionally, never inside a branch
 *-----------------------------------------------------------------------------*)
rtCycle(CLK := bCycleDone);      // 完工沿 / the cycle done edge

(*------------------------------------------------------------------------------
 * 段 1｜错误码与信息位本拍预置（当前周期事实，非锁存）
 *      The error code and the info bit are per scan facts
 *-----------------------------------------------------------------------------*)
uErrorId := TPM_ERR_NONE;        // 预置无错误 / preset no error
_bQtySat := FALSE;               // 信息位复位 / reset the info bit

(*------------------------------------------------------------------------------
 * 段 2｜配置三面闸（电平面，当拍复判，码 01/02）：
 *      目标面（>0 且有限）、平滑系数面（(0,1] 且有限）、窗面（>0）与计时基准面
 *      The three configuration faces, re judged every scan
 *-----------------------------------------------------------------------------*)
_bTgtOk   := (fTaktTargetS > 0.0) AND (fTaktTargetS = fTaktTargetS)
         AND (ABS(fTaktTargetS) <= TPM_FIN_MAX);             // 目标面闸 / the target face gate
_bAlphaOk := (fAlpha > 0.0) AND (fAlpha <= 1.0) AND (fAlpha = fAlpha)
         AND (ABS(fAlpha) <= TPM_FIN_MAX);                   // 平滑系数面闸（(0,1] 域）/ the alpha face gate
_bTimeOk  := (fCallCycleS > 0.0) AND (fCallCycleS = fCallCycleS)
         AND (tEvalWindow > T#0MS);                          // 计时基准面 + 窗面闸（TIME 直接比较）/ the time base and window faces
IF (NOT _bTgtOk) OR (NOT _bTimeOk) THEN
    bError := TRUE;                  // 故障标志（R45 配对，v1.0.1：窗/计时面并入码 01 不再静默）/ the fault flag
    uErrorId := TPM_ERR_TGT;         // 码 01（目标/窗/计时基准面）/ code 01
ELSIF NOT _bAlphaOk THEN
    bError := TRUE;                  // 码 02 / code 02
    uErrorId := TPM_ERR_ALPHA;
ELSE
    bError := FALSE;                 // 配置恢复即清（电平面契约）/ cleared when the configuration recovers
END_IF
IF NOT (_bTgtOk AND _bAlphaOk AND _bTimeOk) THEN
    bValid := FALSE;                 // 任一配置面失效即不出数 / no output while any face fails
    RETURN;                          // 输出全部冻结保持（头注契约）/ all outputs frozen
END_IF
_fWinLimMs := DINT_TO_LREAL(TIME_TO_DINT(tEvalWindow));  // 窗长转毫秒缓存（TIME 本义 ms）[ms] / the window limit in ms

(*------------------------------------------------------------------------------
 * 段 3｜失能相串清账（R 失能清账）：窗累计清零、脉冲基准撤销、bValid 撤销
 *      The disable phase clears the books, the outputs hold frozen
 *-----------------------------------------------------------------------------*)
IF NOT bEnable THEN
    bValid := FALSE;                 // 失能不出数 / no output while disabled
    _bHasPrev := FALSE;              // 撤销脉冲基准（重新使能从下一脉冲起测）/ withdraw the pulse baseline
    _fSinceS := 0.0;                 // 间隔累计清零 / clear the interval accumulator
    _fWinAccMs := 0.0;               // 窗累计清零 / clear the window accumulator
    _uQtyWin := UDINT#0;             // 窗内计数清零 / clear the window count
    _bTaktInit := FALSE;             // EWMA 重新种子（首件语义重置）/ re seed the EWMA
    RETURN;                          // 输出冻结保持 / outputs frozen
END_IF

(*------------------------------------------------------------------------------
 * 段 4｜推进与计件：间隔累计 + 完工沿处理（首件只立基准不出数）
 *      The advance and counting, the first pulse only arms the baseline
 *-----------------------------------------------------------------------------*)
_fSinceS := _fSinceS + fCallCycleS;      // 间隔累计 [s]（推进判据与配置闸不同源）/ accumulate the interval
IF rtCycle.Q THEN                        // 完工沿 / the cycle done edge
    IF _bHasPrev THEN                    // 有基准才出间隔（首件不出数）/ an interval only with a baseline
        fInterval := _fSinceS;           // 取完工间隔 [s] / take the interval
        IF (fInterval <> fInterval) OR (ABS(fInterval) > TPM_FIN_MAX) THEN
            _bQtySat := TRUE;            // 非有限间隔弃用并记信息位（防御，结构性罕见）/ a non finite interval is dropped, marked
        ELSE
            IF NOT _bTaktInit THEN
                fTaktActS := fInterval;  // EWMA 首个有效样本直赋（禁 0 当种子）/ seed the EWMA directly
                _bTaktInit := TRUE;
            ELSE
                fTaktActS := fTaktActS + fAlpha * (fInterval - fTaktActS);  // EWMA 递推 [s] / the EWMA recursion
            END_IF
            bValid := TRUE;              // 首个有效间隔后开始出数 / live after the first valid interval
        END_IF
    ELSE
        bValid := FALSE;                 // 首件前不出数（头注契约）/ no output before the first piece
    END_IF
    _bHasPrev := TRUE;                   // 立脉冲基准 / arm the baseline
    _fSinceS := 0.0;                     // 间隔累计清零 / clear the interval accumulator
    IF _uQtyWin < TPM_U_MAX THEN         // 窗内计数溢出钳位（先闸后加）/ the count saturation clamp
        _uQtyWin := _uQtyWin + UDINT#1;  // 窗内计件 [件] / count the piece in window
    ELSE
        _bQtySat := TRUE;                // 计数饱和记信息位 / mark the saturation
    END_IF
END_IF

(*------------------------------------------------------------------------------
 * 段 5｜评估窗滚动：窗满结算缺口（分母侧显式判：目标面已闸，产量不进分母）
 *      The window roll, the backlog settlement, the quantity never enters a denominator
 *-----------------------------------------------------------------------------*)
_fWinAccMs := _fWinAccMs + fCallCycleS * 1000.0;  // 窗累计 [ms] / accumulate the window
IF _fWinAccMs >= _fWinLimMs THEN         // 窗满滚动判据 / the roll criterion
    fExpectR := (_fWinLimMs / 1000.0) / fTaktTargetS;  // 窗内目标产量 [件]（分母 = 目标，已闸 > 0）/ the expected quantity, the denominator is the gated target
    IF (fExpectR <> fExpectR) OR (fExpectR >= TPM_DINT_MAX) THEN
        _nExpect := TPM_U_MAX;           // 目标产量超 DINT 中转域（v1.0.2 前移至 2^31-1）钳上限 + 信息码（取整前实数上限兜底）/ clamp the expectation to the ceiling
        _bQtySat := TRUE;
    ELSE
        _nExpect := DINT_TO_UDINT(LREAL_TO_DINT(TRUNC(fExpectR)));  // 实数截断为件数（标准转换链，向下取整口径）/ truncate the expectation, standard chain
    END_IF
    IF _nExpect > _uQtyWin THEN
        uQtyBacklog := _nExpect - _uQtyWin;  // 缺口 = 目标 − 实际（无除法面）/ the backlog is the shortfall
    ELSE
        uQtyBacklog := UDINT#0;          // 超产或持平缺口归零（钳位显式）/ no shortfall clamps to zero
    END_IF
    _fWinAccMs := _fWinAccMs - _fWinLimMs;  // 窗基准滚动（保留余量，防长周期漂移）/ roll the window keeping the remainder
    _uQtyWin := UDINT#0;                 // 窗内计数清零 / clear the window count
END_IF

(*------------------------------------------------------------------------------
 * 段 6｜进度偏差与落后判定（分母 = 目标节拍，已闸 > 0；容差判零禁浮点判等）
 *      The pace deviation and the behind verdict, the denominator already gated
 *-----------------------------------------------------------------------------*)
IF bValid THEN                           // 首件前不刷新偏差（输出语义一致）/ no deviation before the first piece
    fPaceDevPct := (fTaktActS - fTaktTargetS) / fTaktTargetS * 100.0;  // 偏差 [%] / the deviation percent
    IF fPaceDevPct > TPM_EPS THEN
        bBehind := TRUE;                 // 正偏差判落后（容差判零）/ a positive deviation means behind
    ELSE
        bBehind := FALSE;                // 非正偏差不落后 / not behind otherwise
    END_IF
END_IF
IF _bQtySat THEN
    uErrorId := TPM_ERR_SAT;             // 信息级码（不置 bError，功能不受影响）/ the info code, no fault flag
END_IF
END_FUNCTION_BLOCK

(* ---- FB_DL_TankAgitationSeq.st ---- *)
(*
  Name        : FB_DL_TankAgitationSeq
  Category    : DL_Process
  Version     : 1.0.0
  Purpose     : 搅拌槽搅拌时序：低速分散 → 高速搅拌 → 维持计时三相编排，液位低禁高速，扭矩过载确认降速回退，转速设定斜坡防冲击；/ Tank agitation sequence: low-speed dispersion, high-speed mixing and hold timing phases, level-low interlock against high speed, torque overload confirmed ramp-down, ramped speed setpoint
  溯源        : 借 isa88 的相语义扩族组织，clean-room 实现
  Boundary    : ① 液位低 → 禁止高速相（联锁），高速已运行则降速回退相；
                ② 扭矩过载判据经确认延时（TON）才降速，瞬时尖峰不误动；
                ③ 三相计时 TON 段 0 无条件刷新 + 相位闸（R40）；
                ④ 降速回退相与故障相分离：回退可恢复（液位/扭矩恢复后重回低速相），组态故障才锁存至复位沿；
                ⑤ 转速设定斜坡逼近防机械冲击；非有限扭矩该拍不判过载（保持当前相）；
                ⑥ 本件为时序编排层，输出转速设定值，不直接驱动变频器（属主边界）。
*)
TYPE E_DL_TasState :
(
    eIdle    := 0,                           (* 未运行（设定转速斜坡回零） / Idle *)
    eLowSpd  := 10,                          (* 低速分散相 / Low-speed dispersion *)
    eHighSpd := 20,                          (* 高速搅拌相 / High-speed mixing *)
    eMaintain:= 30,                          (* 维持计时相 / Hold timing *)
    eRampDn  := 40,                          (* 降速回退相（可恢复，边界④） / Ramp-down recovery *)
    eFault   := 90                           (* 故障锁存相 / Fault latched *)
);
END_TYPE

TYPE E_DL_TasCause :
(
    eNone      := 0,                         (* 无成因 / No cause *)
    eCfgIllegal:= 1,                        (* 组态非法：转速/时长/阈值域越界 / Illegal config *)
    ePhaseBad  := 2                         (* 非法相位兜底 / Illegal phase fallback *)
);
END_TYPE

FUNCTION_BLOCK FB_DL_TankAgitationSeq
VAR_INPUT
    bStart   : BOOL := FALSE;                (* 启动时序命令，上升沿受理 [-] / Start command *)
    bLevelLow: BOOL := FALSE;                (* 液位低信号（联锁源）[-] / Level low signal *)
    fTorque  : REAL := 0.0;                  (* 搅拌扭矩 [%] / Agitator torque *)
    fTqOverLim: REAL := 90.0;                (* 扭矩过载阈，域 > 0 [%] / Torque overload limit *)
    tTqConf  : TIME := T#2S;                 (* 过载确认延时，域 > T#0S [ms] / Overload confirm delay *)
    tLowDwell: TIME := T#60S;                (* 低速分散时长，域 > T#0S [ms] / Low-speed dwell *)
    tHighDwell: TIME := T#300S;              (* 高速搅拌时长 [ms] / High-speed dwell *)
    tMaintain: TIME := T#120S;               (* 维持计时时长 [ms] / Hold duration *)
    fSpdLow  : REAL := 60.0;                 (* 低速设定转速 [rpm] / Low speed setpoint *)
    fSpdHigh : REAL := 180.0;                (* 高速设定转速，域 > 低速 [rpm] / High speed setpoint *)
    fRampRate: REAL := 30.0;                 (* 斜坡率，域 > 0 [rpm/s] / Ramp rate *)
    tScan    : TIME := T#100MS;              (* 扫描周期，域 > T#0S [ms] / Scan period *)
    bEnable  : BOOL := TRUE;                 (* 使能 [-] / Enable *)
    bReset   : BOOL := FALSE;                (* 复位命令，上升沿清故障回空闲 [-] / Reset command *)
END_VAR
VAR_OUTPUT
    fSpdSet  : REAL;                         (* 转速设定出口（斜坡逼近）[rpm] / Ramped speed setpoint outlet *)
    bRunning : BOOL;                         (* 时序运行中指示 [-] / Sequence running indicator *)
    bSeqDone : BOOL;                         (* 时序完成脉冲（单拍）[-] / Sequence done pulse *)
    bRampDn  : BOOL;                         (* 降速回退中指示（状态可查）[-] / Ramp-down indicator *)
    eState   : E_DL_TasState;                (* 状态出口 / State outlet *)
    eCause   : E_DL_TasCause;                (* 成因出口（R190 归因唯一） / Cause outlet *)
    bError   : BOOL;                         (* 故障锁存标志 [-] / Fault latch flag *)
END_VAR
VAR
    _eState : E_DL_TasState := E_DL_TasState.eIdle;  (* 内部相位（CASE 唯一写入目标） / Internal phase *)
    _eCause : E_DL_TasCause := E_DL_TasCause.eNone;  (* 成因锁存量 / Latched cause *)
    rtStart : R_TRIG;                        (* 启动沿实例，段 0 无条件调用 / Start edge instance *)
    rtReset : R_TRIG;                        (* 复位沿实例，段 0 无条件调用 / Reset edge instance *)
    tonLow  : TON;                           (* 低速分散计时（IN 串相位闸，边界③） / Low-speed timer *)
    tonHigh : TON;                           (* 高速搅拌计时（IN 串相位闸） / High-speed timer *)
    tonMaint: TON;                           (* 维持计时（IN 串相位闸） / Hold timer *)
    tonTq   : TON;                           (* 扭矩过载确认计时（IN 串相位 + 有限 + 超限判据，边界②⑤） / Torque confirm timer *)
    _bFault : BOOL;                          (* 故障锁存位 / Latched fault bit *)
    _bCfgBad: BOOL;                          (* 组态非法当拍量 / Illegal config this scan *)
    _bFin   : BOOL;                          (* 扭矩有限性当拍量（边界⑤） / Torque finiteness *)
    _bDoneI : BOOL;                          (* 完成脉冲内部量（统一出口映射，R187） / Done pulse internal *)
    _fTarget: REAL;                          (* 当前相目标转速 [rpm] / Phase target speed *)
    _fStep  : REAL;                          (* 本拍斜坡步长 [rpm] / Ramp step this scan *)
    _fDtSec : REAL;                          (* 扫描周期秒值，域 > eps [s] / Scan period seconds *)
END_VAR
VAR CONSTANT
    DL_TAS_EPS : REAL := 1.0E-6;             (* 判零容差 [-] / Epsilon *)
END_VAR

(* —— 段 0：当拍判据派生 + 实例无条件刷新（R228A；TON 全段 0 无 IF 包裹，边界③） —— *)
_bCfgBad := (fSpdLow <= DL_TAS_EPS) OR (fSpdHigh <= fSpdLow)             (* 转速域闸（高速 > 低速） / Speed gates *)
            OR (fTqOverLim <= DL_TAS_EPS) OR (fRampRate <= DL_TAS_EPS)   (* 阈值/斜率正域闸（边界⑤） / Limit and rate gates *)
            OR NOT (tTqConf > T#0S) OR NOT (tLowDwell > T#0S)            (* 时长域闸（边界③） / Dwell gates *)
            OR NOT (tHighDwell > T#0S) OR NOT (tMaintain > T#0S) OR NOT (tScan > T#0S);   (* 时长域闸续 / Dwell gates cont. *)
rtStart(CLK := bStart);                                  (* 启动沿每拍必调 / Start edge every scan *)
rtReset(CLK := bReset);                                  (* 复位沿每拍必调 / Reset edge every scan *)
_bFin := (fTorque = fTorque) AND ((fTorque - fTorque) = (fTorque - fTorque));   (* 扭矩 NaN 自反 + Inf 差判闸（边界⑤） / Torque NaN and Inf gate *)
_fDtSec := TIME_TO_LREAL(tScan) / 1000.0;                (* 扫描周期秒化（除子常量 1000） / Scan period seconds *)
_fStep := fRampRate * _fDtSec;                           (* 斜坡步长 = 率 × 周期秒值（边界⑤） / Ramp step *)
tonLow(IN := (_eState = E_DL_TasState.eLowSpd), PT := tLowDwell);        (* 低速计时：相位闸 + 无条件调用（R40） / Low timer *)
tonHigh(IN := (_eState = E_DL_TasState.eHighSpd), PT := tHighDwell);     (* 高速计时：相位闸 + 无条件调用 / High timer *)
tonMaint(IN := (_eState = E_DL_TasState.eMaintain), PT := tMaintain);    (* 维持计时：相位闸 + 无条件调用 / Hold timer *)
tonTq(IN := (_eState = E_DL_TasState.eHighSpd) AND _bFin AND (fTorque > fTqOverLim), PT := tTqConf);   (* 过载确认：相闸 + 有限闸 + 超限直比（边界②⑤） / Torque confirm *)

(* —— 段 1：单拍量预清零（R107） —— *)
_bDoneI := FALSE;                                        (* 完成脉冲内部量预清 / Done preset *)
bSeqDone := FALSE;                                       (* 完成脉冲出口预清 / Done outlet preset *)
bRunning := FALSE;                                       (* 运行指示出口预清（派生拍覆盖） / Running preset *)
bRampDn := FALSE;                                        (* 回退指示出口预清 / Ramp-down preset *)

(* —— 段 2：复位沿处理（作用域：清故障 + 回空闲 + 设定归零，R283 逐项声明） —— *)
IF rtReset.Q THEN
    _bFault := FALSE;                                    (* 清故障锁存 / Clear fault *)
    _eCause := E_DL_TasCause.eNone;                      (* 清成因 / Clear cause *)
    _eState := E_DL_TasState.eIdle;                      (* 回空闲相 / Back to idle *)
END_IF

(* —— 段 3：组态故障锁存（锁存至复位沿，R189） —— *)
IF _bCfgBad AND NOT _bFault THEN
    _bFault := TRUE;                                     (* 锁存故障位 / Latch fault *)
    _eCause := E_DL_TasCause.eCfgIllegal;                (* 成因：组态非法 / Cause illegal config *)
    _eState := E_DL_TasState.eFault;                     (* 同步迁故障相 / Migrate to fault *)
END_IF

(* —— 段 4：CASE 主状态机（ELSE 兜底迁 eFault，红线 6） —— *)
CASE _eState OF
    E_DL_TasState.eIdle:                                 (* 空闲：目标转速 0（斜坡归零防冲击，边界⑤） / Idle *)
        _fTarget := 0.0;                                 (* 目标转速零 / Target zero *)
        IF rtStart.Q AND bEnable AND NOT _bFault AND NOT bLevelLow THEN   (* 启动受理：液位低禁进入（联锁前置，边界①） / Start gating *)
            _eState := E_DL_TasState.eLowSpd;            (* 进入低速分散相 / Enter low-speed *)
        END_IF
    E_DL_TasState.eLowSpd:                               (* 低速分散相：计时满且液位不低 → 高速 / Low-speed *)
        _fTarget := fSpdLow;                             (* 目标 = 低速设定 / Target low speed *)
        bRunning := TRUE;                                (* 运行指示出口 / Running indicator *)
        IF NOT bEnable THEN
            _eState := E_DL_TasState.eIdle;              (* 失能回空闲 / Back to idle *)
        ELSIF tonLow.Q AND NOT bLevelLow THEN            (* 计时满 + 液位不低才进高速（联锁，边界①） / Dwell done and level ok *)
            _eState := E_DL_TasState.eHighSpd;           (* 进入高速搅拌相 / Enter high-speed *)
        END_IF
    E_DL_TasState.eHighSpd:                              (* 高速搅拌相：液位低/过载回退，计时满 → 维持 / High-speed *)
        _fTarget := fSpdHigh;                            (* 目标 = 高速设定 / Target high speed *)
        bRunning := TRUE;                                (* 运行指示出口 / Running indicator *)
        IF NOT bEnable THEN
            _eState := E_DL_TasState.eIdle;              (* 失能回空闲 / Back to idle *)
        ELSIF bLevelLow OR tonTq.Q THEN                  (* 液位低（边界①）或过载确认（边界②）：降速回退 / Level low or overload confirmed *)
            _eState := E_DL_TasState.eRampDn;            (* 进降速回退相（可恢复，边界④） / Enter ramp-down *)
        ELSIF tonHigh.Q THEN
            _eState := E_DL_TasState.eMaintain;          (* 计时满进维持相 / Enter hold *)
        END_IF
    E_DL_TasState.eMaintain:                             (* 维持计时相：低速维持 + 计时满完成 / Hold *)
        _fTarget := fSpdLow;                             (* 维持相目标 = 低速 / Target low speed *)
        bRunning := TRUE;                                (* 运行指示出口 / Running indicator *)
        IF NOT bEnable THEN
            _eState := E_DL_TasState.eIdle;              (* 失能回空闲 / Back to idle *)
        ELSIF tonMaint.Q THEN
            _bDoneI := TRUE;                             (* 时序完成内部置位（R187） / Done internal *)
            _eState := E_DL_TasState.eIdle;              (* 回空闲（设定斜坡归零） / Back to idle *)
        END_IF
    E_DL_TasState.eRampDn:                               (* 降速回退相：斜坡到低速 → 重回低速相（可恢复，边界④） / Ramp-down *)
        _fTarget := fSpdLow;                             (* 回退目标 = 低速 / Target low speed *)
        bRunning := TRUE;                                (* 回退仍属运行（状态可查） / Running indicator *)
        bRampDn := TRUE;                                 (* 回退指示出口 / Ramp-down indicator *)
        IF NOT bEnable THEN
            _eState := E_DL_TasState.eIdle;              (* 失能回空闲 / Back to idle *)
        ELSIF ABS(fSpdSet - fSpdLow) <= _fStep THEN      (* 斜坡到位（容差直比，非浮点等值） / Ramp arrived *)
            _eState := E_DL_TasState.eLowSpd;            (* 重回低速分散相（恢复，边界④） / Back to low-speed *)
        END_IF
    E_DL_TasState.eFault:                                (* 故障相：冻结保持，仅复位沿出 / Fault *)
        _fTarget := 0.0;                                 (* 故障相目标归零（安全侧确定值） / Target zero in fault *)
        ;                                                (* 锁存回放（R28） / Replay from latch *)
    ELSE                                                 (* 非法相位兜底迁安全态 / Illegal phase fallback *)
        _eState := E_DL_TasState.eFault; _bFault := TRUE;    (* 迁故障相 + 同步锁存 / To fault and latch *)
        _eCause := E_DL_TasCause.ePhaseBad;              (* 成因：非法相位 / Cause illegal phase *)
END_CASE

(* —— 段 4B：设定斜坡逼近（防机械冲击，边界⑤；容差直比防浮点等值抖动） —— *)
IF fSpdSet < (_fTarget - _fStep) THEN
    fSpdSet := fSpdSet + _fStep;                         (* 正向斜坡步进 / Ramp up *)
ELSIF fSpdSet > (_fTarget + _fStep) THEN
    fSpdSet := fSpdSet - _fStep;                         (* 负向斜坡步进 / Ramp down *)
ELSE
    fSpdSet := _fTarget;                                 (* 步长内直达目标 / Reach target *)
END_IF

(* —— 段 5：出口映射（内部 _b* → 输出单拍，R187；bError/eState 同源，R191） —— *)
bSeqDone := _bDoneI;                                     (* 完成脉冲单拍出口 / Done pulse outlet *)
bError := _bFault;                                       (* 故障标志镜像 / Fault flag mirror *)
eState := _eState;                                       (* 状态出口 / State outlet *)
eCause := _eCause;                                       (* 成因出口 / Cause outlet *)
END_FUNCTION_BLOCK
